screen "Visu_ES_rep5_6" 1280x800, template "Modèle_ES"
   GraphicView "Vue de graphique_1" at 62,186 size 76x151; Picture "Graphique_4"
   TextField "Champ de texte_1" at 43,144 size 59x25; Text 'REP 5'
   Rectangle "Rectangle_2" at 189,244 size 20x20
      Appearance <- "I_det_photo_02"
   TextField "Champ de texte_2" at 215,242 size 136x25; Text 'Det. Photo. 5'
   Rectangle "Rectangle_3" at 189,266 size 20x20
      Appearance <- "AlwaysFALSE"
   TextField "Champ de texte_3" at 215,264 size 53x25; Text 'Libre'
   Rectangle "Rectangle_4" at 189,288 size 20x20
      Appearance <- "AlwaysFALSE"
   TextField "Champ de texte_4" at 215,286 size 53x25; Text 'Libre'
   Rectangle "Rectangle_5" at 189,310 size 20x20
      Appearance <- "AlwaysFALSE"
   TextField "Champ de texte_5" at 215,308 size 53x25; Text 'Libre'
   Rectangle "Rectangle_6" at 189,332 size 20x20
      Appearance <- "AlwaysFALSE"
   TextField "Champ de texte_6" at 215,330 size 53x25; Text 'Libre'
   Rectangle "Rectangle_7" at 189,354 size 20x20
      Appearance <- "AlwaysFALSE"
   TextField "Champ de texte_7" at 215,352 size 53x25; Text 'Libre'
   Rectangle "Rectangle_8" at 189,376 size 20x20
      Appearance <- "AlwaysFALSE"
   TextField "Champ de texte_8" at 215,374 size 53x25; Text 'Libre'
   Rectangle "Rectangle_9" at 189,398 size 20x20
      Appearance <- "AlwaysFALSE"
   TextField "Champ de texte_9" at 215,396 size 53x25; Text 'Libre'
   Rectangle "Rectangle_10" at 399,244 size 20x20
      Appearance <- "I_det_photo_01"
   TextField "Champ de texte_10" at 425,242 size 136x25; Text 'Det. Photo. 4'
   Rectangle "Rectangle_11" at 399,266 size 20x20
      Appearance <- "I_det_photo_03"
   TextField "Champ de texte_11" at 425,264 size 136x25; Text 'Det. Photo. 6'
   Rectangle "Rectangle_12" at 399,288 size 20x20
      Appearance <- "AlwaysFALSE"
   TextField "Champ de texte_12" at 425,286 size 53x25; Text 'Libre'
   Rectangle "Rectangle_13" at 399,310 size 20x20
      Appearance <- "I_libre_I23"
   TextField "Champ de texte_13" at 425,308 size 53x25; Text 'Libre'
   Rectangle "Rectangle_14" at 399,332 size 20x20
      Appearance <- "AlwaysFALSE"
   TextField "Champ de texte_14" at 425,330 size 53x25; Text 'Libre'
   Rectangle "Rectangle_15" at 399,354 size 20x20
      Appearance <- "AlwaysFALSE"
   TextField "Champ de texte_15" at 425,352 size 53x25; Text 'Libre'
   Rectangle "Rectangle_16" at 399,376 size 20x20
      Appearance <- "AlwaysFALSE"
   TextField "Champ de texte_16" at 425,374 size 53x25; Text 'Libre'
   Rectangle "Rectangle_17" at 399,398 size 20x20
      Appearance <- "AlwaysFALSE"
   TextField "Champ de texte_17" at 425,396 size 53x25; Text 'Libre'
   TextField "Champ de texte_34" at 170,173 size 459x25; Text 'ENTREES'
   TextField "Champ de texte_35" at 189,219 size 59x25; Text '%I12'
   TextField "Champ de texte_37" at 399,219 size 59x25; Text '%I13'
   GraphicView "Vue de graphique_2" at 62,454 size 76x151; Picture "Graphique_4"
   TextField "Champ de texte_18" at 43,412 size 59x25; Text 'REP 6'
   Rectangle "Rectangle_20" at 189,512 size 20x20
      Appearance <- "I_Det_Photo_8"
   TextField "Champ de texte_19" at 215,510 size 130x25; Text 'Det. Photo. 8'
   Rectangle "Rectangle_21" at 189,534 size 20x20
      Appearance <- "AlwaysFALSE"
   TextField "Champ de texte_20" at 215,532 size 53x25; Text 'Libre'
   Rectangle "Rectangle_22" at 189,556 size 20x20
      Appearance <- "AlwaysFALSE"
   TextField "Champ de texte_21" at 215,554 size 53x25; Text 'Libre'
   Rectangle "Rectangle_23" at 189,578 size 20x20
      Appearance <- "AlwaysFALSE"
   TextField "Champ de texte_22" at 215,576 size 53x25; Text 'Libre'
   Rectangle "Rectangle_24" at 189,600 size 20x20
      Appearance <- "AlwaysFALSE"
   TextField "Champ de texte_23" at 215,598 size 53x25; Text 'Libre'
   Rectangle "Rectangle_25" at 189,622 size 20x20
      Appearance <- "AlwaysFALSE"
   TextField "Champ de texte_24" at 215,620 size 53x25; Text 'Libre'
   Rectangle "Rectangle_26" at 189,644 size 20x20
      Appearance <- "AlwaysFALSE"
   TextField "Champ de texte_25" at 215,642 size 53x25; Text 'Libre'
   Rectangle "Rectangle_27" at 189,666 size 20x20
      Appearance <- "AlwaysFALSE"
   TextField "Champ de texte_26" at 215,664 size 53x25; Text 'Libre'
   Rectangle "Rectangle_28" at 399,512 size 20x20
      Appearance <- "I_Det_Photo_7"
   TextField "Champ de texte_27" at 425,510 size 130x25; Text 'Det. Photo. 7'
   Rectangle "Rectangle_29" at 399,534 size 20x20
      Appearance <- "I_Det_Photo_9"
   TextField "Champ de texte_28" at 425,532 size 130x25; Text 'Det. Photo. 9'
   Rectangle "Rectangle_30" at 399,556 size 20x20
      Appearance <- "AlwaysFALSE"
   TextField "Champ de texte_29" at 425,554 size 53x25; Text 'Libre'
   Rectangle "Rectangle_31" at 399,578 size 20x20
      Appearance <- "AlwaysFALSE"
   TextField "Champ de texte_30" at 425,576 size 53x25; Text 'Libre'
   Rectangle "Rectangle_32" at 399,600 size 20x20
      Appearance <- "AlwaysFALSE"
   TextField "Champ de texte_31" at 425,598 size 53x25; Text 'Libre'
   Rectangle "Rectangle_34" at 399,622 size 20x20
      Appearance <- "AlwaysFALSE"
   TextField "Champ de texte_32" at 425,620 size 53x25; Text 'Libre'
   Rectangle "Rectangle_36" at 399,644 size 20x20
      Appearance <- "AlwaysFALSE"
   TextField "Champ de texte_33" at 425,642 size 53x25; Text 'Libre'
   Rectangle "Rectangle_37" at 399,666 size 20x20
      Appearance <- "AlwaysFALSE"
   TextField "Champ de texte_36" at 425,664 size 53x25; Text 'Libre'
   TextField "Champ de texte_38" at 170,441 size 459x25; Text 'ENTREES'
   TextField "Champ de texte_39" at 189,487 size 59x25; Text '%I14'
   TextField "Champ de texte_40" at 399,487 size 59x25; Text '%I15'

screen "Visu_ES_Ilot01" 1280x800, template "Modèle_ES"
   TextField "Champ de texte_1" at 43,144 size 80x25; Text 'ILOT 01'
   Rectangle "Rectangle_2" at 273,244 size 20x20
      Appearance <- "O_Rentrer_Butée_01"
   TextField "Champ de texte_2" at 299,242 size 167x25; Text 'Rentrer Butée 01'
   Rectangle "Rectangle_3" at 273,266 size 20x20
      Appearance <- "O_Rentrer_Butée_EL_01"
   TextField "Champ de texte_3" at 299,264 size 202x25; Text 'Rentrer But. Elev. 01'
   Rectangle "Rectangle_4" at 273,288 size 20x20
      Appearance <- "O_Monter_EL_01"
   TextField "Champ de texte_4" at 299,286 size 184x25; Text 'Sortir Elevateur 01'
   Rectangle "Rectangle_5" at 273,310 size 20x20
      Appearance <- "O_Desc_EL_01"
   TextField "Champ de texte_5" at 299,308 size 201x25; Text 'Rentrer Elevateur 01'
   Rectangle "Rectangle_6" at 273,332 size 20x20
      Appearance <- "O_Rentrer_Butée_02"
   TextField "Champ de texte_6" at 299,330 size 167x25; Text 'Rentrer Butée 02'
   Rectangle "Rectangle_7" at 273,354 size 20x20
      Appearance <- "O_Rentrer_Butée_EL_02"
   TextField "Champ de texte_7" at 299,352 size 202x25; Text 'Rentrer But. Elev. 02'
   Rectangle "Rectangle_8" at 273,376 size 20x20
      Appearance <- "O_Monter_EL_02"
   TextField "Champ de texte_8" at 299,374 size 184x25; Text 'Sortir Elevateur 02'
   Rectangle "Rectangle_9" at 273,398 size 20x20
      Appearance <- "O_Desc_EL_02"
   TextField "Champ de texte_9" at 299,396 size 201x25; Text 'Rentrer Elevateur 02'
   Rectangle "Rectangle_10" at 483,244 size 20x20
      Appearance <- "O_Rentrer_Butée_03"
   TextField "Champ de texte_10" at 509,242 size 167x25; Text 'Rentrer Butée 03'
   Rectangle "Rectangle_11" at 483,266 size 20x20
      Appearance <- "O_Rentrer_Butée_EL_03"
   TextField "Champ de texte_11" at 509,264 size 202x25; Text 'Rentrer But. Elev. 03'
   Rectangle "Rectangle_12" at 483,288 size 20x20
      Appearance <- "O_Monter_EL_03"
   TextField "Champ de texte_12" at 509,286 size 184x25; Text 'Sortir Elevateur 03'
   Rectangle "Rectangle_13" at 483,310 size 20x20
      Appearance <- "O_Desc_EL_03"
   TextField "Champ de texte_13" at 509,308 size 201x25; Text 'Rentrer Elevateur 03'
   Rectangle "Rectangle_14" at 483,332 size 20x20
      Appearance <- "O_Rentrer_Butée_04"
   TextField "Champ de texte_14" at 509,330 size 167x25; Text 'Rentrer Butée 04'
   Rectangle "Rectangle_15" at 483,354 size 20x20
      Appearance <- "O_Rentrer_Butée_EL_04"
   TextField "Champ de texte_15" at 509,352 size 202x25; Text 'Rentrer But. Elev. 04'
   Rectangle "Rectangle_16" at 483,376 size 20x20
      Appearance <- "O_Monter_EL_04"
   TextField "Champ de texte_16" at 509,374 size 184x25; Text 'Sortir Elevateur 04'
   Rectangle "Rectangle_17" at 483,398 size 20x20
      Appearance <- "O_Desc_EL_04"
   TextField "Champ de texte_17" at 509,396 size 201x25; Text 'Rentrer Elevateur 04'
   TextField "Champ de texte_34" at 254,173 size 880x25; Text 'SORTIES'
   TextField "Champ de texte_35" at 273,219 size 64x25; Text '%Q10'
   TextField "Champ de texte_37" at 483,219 size 64x25; Text '%Q11'
   GraphicView "Vue de graphique_3" at 58,184 size 154x109; Picture "Graphique_5"
   Rectangle "Rectangle_18" at 692,244 size 20x20
      Appearance <- "O_Rentrer_Butée_05"
   TextField "Champ de texte_18" at 718,242 size 167x25; Text 'Rentrer Butée 05'
   Rectangle "Rectangle_19" at 692,266 size 20x20
      Appearance <- "O_Rentrer_Butée_EL_05"
   TextField "Champ de texte_19" at 718,264 size 202x25; Text 'Rentrer But. Elev. 05'
   Rectangle "Rectangle_20" at 692,288 size 20x20
      Appearance <- "O_Monter_EL_05"
   TextField "Champ de texte_20" at 718,286 size 184x25; Text 'Sortir Elevateur 05'
   Rectangle "Rectangle_21" at 692,310 size 20x20
      Appearance <- "O_Desc_EL_05"
   TextField "Champ de texte_21" at 718,308 size 201x25; Text 'Rentrer Elevateur 05'
   Rectangle "Rectangle_22" at 692,332 size 20x20
      Appearance <- "O_Rentrer_Butée_06"
   TextField "Champ de texte_22" at 718,330 size 167x25; Text 'Rentrer Butée 06'
   Rectangle "Rectangle_23" at 692,354 size 20x20
      Appearance <- "O_Rentrer_Butée_EL_06"
   TextField "Champ de texte_23" at 718,352 size 202x25; Text 'Rentrer But. Elev. 06'
   Rectangle "Rectangle_24" at 692,376 size 20x20
      Appearance <- "O_Monter_EL_06"
   TextField "Champ de texte_24" at 718,374 size 184x25; Text 'Sortir Elevateur 06'
   Rectangle "Rectangle_25" at 692,398 size 20x20
      Appearance <- "O_Desc_EL_06"
   TextField "Champ de texte_25" at 718,396 size 201x25; Text 'Rentrer Elevateur 06'
   Rectangle "Rectangle_26" at 902,244 size 20x20
      Appearance <- "O_Rentrer_Butée_07"
   TextField "Champ de texte_26" at 928,242 size 167x25; Text 'Rentrer Butée 07'
   Rectangle "Rectangle_27" at 902,266 size 20x20
      Appearance <- "O_Rentrer_Butée_EL_07"
   TextField "Champ de texte_27" at 928,264 size 202x25; Text 'Rentrer But. Elev. 07'
   Rectangle "Rectangle_28" at 902,288 size 20x20
      Appearance <- "O_Monter_EL_07"
   TextField "Champ de texte_28" at 928,286 size 184x25; Text 'Sortir Elevateur 07'
   Rectangle "Rectangle_29" at 902,310 size 20x20
      Appearance <- "O_Desc_EL_07"
   TextField "Champ de texte_29" at 928,308 size 201x25; Text 'Rentrer Elevateur 07'
   Rectangle "Rectangle_30" at 902,332 size 20x20
      Appearance <- "O_Op_Porte_Vision"
   TextField "Champ de texte_30" at 928,330 size 185x25; Text 'Ouvrir Porte Vision'
   Rectangle "Rectangle_31" at 902,354 size 20x20
      Appearance <- "O_Cl_porte_Vision"
   TextField "Champ de texte_31" at 928,352 size 192x25; Text 'Fermer Porte Vision'
   Rectangle "Rectangle_32" at 902,376 size 20x20
      Appearance <- "I_libre_I26"
   TextField "Champ de texte_32" at 928,374 size 53x25; Text 'Libre'
   Rectangle "Rectangle_34" at 902,398 size 20x20
      Appearance <- "I_libre_I27"
   TextField "Champ de texte_33" at 928,396 size 53x25; Text 'Libre'
   TextField "Champ de texte_36" at 692,219 size 64x25; Text '%Q12'
   TextField "Champ de texte_38" at 902,219 size 64x25; Text '%Q13'

screen "Visu_ES_Ilot02" 1280x800, template "Modèle_ES"
   TextField "Champ de texte_1" at 43,144 size 80x25; Text 'ILOT 02'
   Rectangle "Rectangle_2" at 273,244 size 20x20
      Appearance <- "O_Sortir_Blocage_boite_01"
   TextField "Champ de texte_2" at 299,242 size 184x25; Text 'Sortir Verin 1 bloc.'
   Rectangle "Rectangle_3" at 273,266 size 20x20
      Appearance <- "O_Rentrer_Blocage_boite_01"
   TextField "Champ de texte_3" at 299,264 size 201x25; Text 'Rentrer Verin 1 bloc.'
   Rectangle "Rectangle_4" at 273,288 size 20x20
      Appearance <- "O_Sortir_Blocage_boite_02"
   TextField "Champ de texte_4" at 299,286 size 184x25; Text 'Sortir Verin 2 bloc.'
   Rectangle "Rectangle_5" at 273,310 size 20x20
      Appearance <- "O_Rentrer_Blocage_boite_02"
   TextField "Champ de texte_5" at 299,308 size 201x25; Text 'Rentrer Verin 2 bloc.'
   Rectangle "Rectangle_6" at 273,332 size 20x20
      Appearance <- "O_Sortir_Blocage_boite_03"
   TextField "Champ de texte_6" at 299,330 size 184x25; Text 'Sortir Verin 3 bloc.'
   Rectangle "Rectangle_7" at 273,354 size 20x20
      Appearance <- "O_Rentrer_Blocage_boite_03"
   TextField "Champ de texte_7" at 299,352 size 201x25; Text 'Rentrer Verin 3 bloc.'
   Rectangle "Rectangle_8" at 273,376 size 20x20
      Appearance <- "O_Sortir_Blocage_boite_04"
   TextField "Champ de texte_8" at 299,374 size 184x25; Text 'Sortir Verin 4 bloc.'
   Rectangle "Rectangle_9" at 273,398 size 20x20
      Appearance <- "O_Rentrer_Blocage_boite_04"
   TextField "Champ de texte_9" at 299,396 size 201x25; Text 'Rentrer Verin 4 bloc.'
   Rectangle "Rectangle_10" at 483,244 size 20x20
      Appearance <- "I_libre_I20"
   TextField "Champ de texte_10" at 509,242 size 53x25; Text 'Libre'
   Rectangle "Rectangle_11" at 483,266 size 20x20
      Appearance <- "I_libre_I21"
   TextField "Champ de texte_11" at 509,264 size 53x25; Text 'Libre'
   Rectangle "Rectangle_12" at 483,288 size 20x20
      Appearance <- "I_libre_I22"
   TextField "Champ de texte_12" at 509,286 size 53x25; Text 'Libre'
   Rectangle "Rectangle_13" at 483,310 size 20x20
      Appearance <- "I_libre_I23"
   TextField "Champ de texte_13" at 509,308 size 53x25; Text 'Libre'
   Rectangle "Rectangle_14" at 483,332 size 20x20
      Appearance <- "I_libre_I24"
   TextField "Champ de texte_14" at 509,330 size 53x25; Text 'Libre'
   Rectangle "Rectangle_15" at 483,354 size 20x20
      Appearance <- "I_libre_I25"
   TextField "Champ de texte_15" at 509,352 size 53x25; Text 'Libre'
   Rectangle "Rectangle_16" at 483,376 size 20x20
      Appearance <- "I_libre_I26"
   TextField "Champ de texte_16" at 509,374 size 53x25; Text 'Libre'
   Rectangle "Rectangle_17" at 483,398 size 20x20
      Appearance <- "I_libre_I27"
   TextField "Champ de texte_17" at 509,396 size 53x25; Text 'Libre'
   TextField "Champ de texte_34" at 254,173 size 880x25; Text 'SORTIES'
   TextField "Champ de texte_35" at 273,219 size 64x25; Text '%Q14'
   TextField "Champ de texte_37" at 483,219 size 64x25; Text '%Q15'
   GraphicView "Vue de graphique_3" at 58,184 size 154x109; Picture "Graphique_5"
   Rectangle "Rectangle_18" at 692,244 size 20x20
      Appearance <- "I_En_Service"
   TextField "Champ de texte_18" at 718,242 size 53x25; Text 'Libre'
   Rectangle "Rectangle_19" at 692,266 size 20x20
      Appearance <- "I_En_Arret_Urgence"
   TextField "Champ de texte_19" at 718,264 size 53x25; Text 'Libre'
   Rectangle "Rectangle_20" at 692,288 size 20x20
      Appearance <- "I_En_Manuel"
   TextField "Champ de texte_20" at 718,286 size 53x25; Text 'Libre'
   Rectangle "Rectangle_21" at 692,310 size 20x20
      Appearance <- "I_En_Automatique"
   TextField "Champ de texte_21" at 718,308 size 53x25; Text 'Libre'
   Rectangle "Rectangle_22" at 692,332 size 20x20
      Appearance <- "I_porte_non_réarmée"
   TextField "Champ de texte_22" at 718,330 size 53x25; Text 'Libre'
   Rectangle "Rectangle_23" at 692,354 size 20x20
      Appearance <- "I_porte_01_Op"
   TextField "Champ de texte_23" at 718,352 size 53x25; Text 'Libre'
   Rectangle "Rectangle_24" at 692,376 size 20x20
      Appearance <- "I_porte_02_Op"
   TextField "Champ de texte_24" at 718,374 size 53x25; Text 'Libre'
   Rectangle "Rectangle_25" at 692,398 size 20x20
      Appearance <- "I_libre_I07"
   TextField "Champ de texte_25" at 718,396 size 53x25; Text 'Libre'
   Rectangle "Rectangle_26" at 902,244 size 20x20
      Appearance <- "I_libre_I20"
   TextField "Champ de texte_26" at 928,242 size 53x25; Text 'Libre'
   Rectangle "Rectangle_27" at 902,266 size 20x20
      Appearance <- "I_libre_I21"
   TextField "Champ de texte_27" at 928,264 size 53x25; Text 'Libre'
   Rectangle "Rectangle_28" at 902,288 size 20x20
      Appearance <- "I_libre_I22"
   TextField "Champ de texte_28" at 928,286 size 53x25; Text 'Libre'
   Rectangle "Rectangle_29" at 902,310 size 20x20
      Appearance <- "I_libre_I23"
   TextField "Champ de texte_29" at 928,308 size 53x25; Text 'Libre'
   Rectangle "Rectangle_30" at 902,332 size 20x20
      Appearance <- "I_libre_I24"
   TextField "Champ de texte_30" at 928,330 size 53x25; Text 'Libre'
   Rectangle "Rectangle_31" at 902,354 size 20x20
      Appearance <- "I_libre_I25"
   TextField "Champ de texte_31" at 928,352 size 53x25; Text 'Libre'
   Rectangle "Rectangle_32" at 902,376 size 20x20
      Appearance <- "I_libre_I26"
   TextField "Champ de texte_32" at 928,374 size 53x25; Text 'Libre'
   Rectangle "Rectangle_34" at 902,398 size 20x20
      Appearance <- "I_libre_I27"
   TextField "Champ de texte_33" at 928,396 size 53x25; Text 'Libre'
   TextField "Champ de texte_36" at 692,219 size 64x25; Text '%Q16'
   TextField "Champ de texte_38" at 902,219 size 64x25; Text '%Q17'

screen "Mode_Manuel_B01" 1280x800, template "Modèle_Manu"
   TextField "Champ de texte_34" at 33,135 size 584x25; Text 'Hyppodrome Poste 01'
   Button "Bouton_1" at 39,179 size 169x68; TextOff 'MONTER BUTEE'
      on Press: SetBit("Touche_Tch_Manu{0}")
      on Release: ResetBit("Touche_Tch_Manu{0}")
      Appearance <- "O_Rentrer_Butée_01"
   Button "Bouton_2" at 39,255 size 169x68; TextOff 'DESCENDRE BUTEE'
      on Press: SetBit("Touche_Tch_Manu{1}")
      on Release: ResetBit("Touche_Tch_Manu{1}")
   Button "Bouton_3" at 220,179 size 169x68; TextOff 'MONTER BUTEE ELEVATEUR'
      on Press: SetBit("Touche_Tch_Manu{2}")
      on Release: ResetBit("Touche_Tch_Manu{2}")
   Button "Bouton_4" at 220,255 size 169x68; TextOff 'DESCENDRE BUTEE ELEVATEUR'
      on Press: SetBit("Touche_Tch_Manu{3}")
      on Release: ResetBit("Touche_Tch_Manu{3}")
   Button "Bouton_5" at 39,331 size 169x68; TextOff 'MONTER ELEVATEUR'
      on Press: SetBit("Touche_Tch_Manu{4}")
      on Release: ResetBit("Touche_Tch_Manu{4}")
   Button "Bouton_6" at 220,331 size 169x68; TextOff 'DESCENDRE ELEVATEUR'
      on Press: SetBit("Touche_Tch_Manu{5}")
      on Release: ResetBit("Touche_Tch_Manu{5}")
   Rectangle "Rectangle_2" at 404,181 size 20x20
      Appearance <- "I_Pres_Pal_B01"
   TextField "Champ de texte_2" at 430,179 size 168x25; Text 'Presence pal B01'
   Rectangle "Rectangle_3" at 404,203 size 20x20
      Appearance <- "I_Pres_Elev_B01"
   TextField "Champ de texte_3" at 430,201 size 178x25; Text 'Presence Elev B01'
   Rectangle "Rectangle_4" at 404,225 size 20x20
      Appearance <- "I_Elev_01_Bas"
   TextField "Champ de texte_4" at 430,223 size 177x25; Text 'Elevateur Bas B01'
   Rectangle "Rectangle_5" at 404,247 size 20x20
      Appearance <- "I_Elev_01_Haut"
   TextField "Champ de texte_5" at 430,245 size 188x25; Text 'Elevateur Haut B01'
   TextField "Champ de texte_1" at 34,419 size 584x25; Text 'Hyppodrome Poste 02'
   Button "Bouton_7" at 38,460 size 169x68; TextOff 'MONTER BUTEE'
      on Release: ResetBit("Touche_Tch_Manu{6}")
      on Press: SetBit("Touche_Tch_Manu{6}")
   Button "Bouton_8" at 38,536 size 169x68; TextOff 'DESCENDRE BUTEE'
      on Release: ResetBit("Touche_Tch_Manu{7}")
      on Press: SetBit("Touche_Tch_Manu{7}")
   Button "Bouton_9" at 219,460 size 169x68; TextOff 'MONTER BUTEE ELEVATEUR'
      on Release: ResetBit("Touche_Tch_Manu{8}")
      on Press: SetBit("Touche_Tch_Manu{8}")
   Button "Bouton_10" at 219,536 size 169x68; TextOff 'DESCENDRE BUTEE ELEVATEUR'
      on Release: ResetBit("Touche_Tch_Manu{9}")
      on Press: SetBit("Touche_Tch_Manu{9}")
   Button "Bouton_11" at 38,612 size 169x68; TextOff 'MONTER ELEVATEUR'
      on Release: ResetBit("Touche_Tch_Manu{10}")
      on Press: SetBit("Touche_Tch_Manu{10}")
   Button "Bouton_12" at 219,612 size 169x68; TextOff 'DESCENDRE ELEVATEUR'
      on Release: ResetBit("Touche_Tch_Manu{11}")
      on Press: SetBit("Touche_Tch_Manu{11}")
   Rectangle "Rectangle_7" at 403,462 size 20x20
      Appearance <- "I_Pres_Pal_B02"
   TextField "Champ de texte_6" at 429,460 size 168x25; Text 'Presence pal B02'
   Rectangle "Rectangle_8" at 403,484 size 20x20
      Appearance <- "I_Pres_Elev_B02"
   TextField "Champ de texte_7" at 429,482 size 178x25; Text 'Presence Elev B02'
   Rectangle "Rectangle_9" at 403,506 size 20x20
      Appearance <- "I_Elev_02_Bas"
   TextField "Champ de texte_8" at 429,504 size 177x25; Text 'Elevateur Bas B02'
   Rectangle "Rectangle_10" at 403,528 size 20x20
      Appearance <- "I_Elev_02_Haut"
   TextField "Champ de texte_9" at 429,526 size 188x25; Text 'Elevateur Haut B02'
   TextField "Champ de texte_10" at 665,138 size 584x25; Text 'Hyppodrome Poste 03'
   Button "Bouton_13" at 669,179 size 169x68; TextOff 'MONTER BUTEE'
      on Release: ResetBit("Touche_Tch_Manu{12}")
      on Press: SetBit("Touche_Tch_Manu{12}")
   Button "Bouton_14" at 669,255 size 169x68; TextOff 'DESCENDRE BUTEE'
      on Release: ResetBit("Touche_Tch_Manu{13}")
      on Press: SetBit("Touche_Tch_Manu{13}")
   Button "Bouton_15" at 850,179 size 169x68; TextOff 'MONTER BUTEE ELEVATEUR'
      on Release: ResetBit("Touche_Tch_Manu{14}")
      on Press: SetBit("Touche_Tch_Manu{14}")
   Button "Bouton_16" at 850,255 size 169x68; TextOff 'DESCENDRE BUTEE ELEVATEUR'
      on Release: ResetBit("Touche_Tch_Manu{15}")
      on Press: SetBit("Touche_Tch_Manu{15}")
   Button "Bouton_17" at 669,331 size 169x68; TextOff 'MONTER ELEVATEUR'
      on Release: ResetBit("Touche_Tch_Manu{16}")
      on Press: SetBit("Touche_Tch_Manu{16}")
   Button "Bouton_18" at 850,331 size 169x68; TextOff 'DESCENDRE ELEVATEUR'
      on Release: ResetBit("Touche_Tch_Manu{17}")
      on Press: SetBit("Touche_Tch_Manu{17}")
   Rectangle "Rectangle_13" at 1034,181 size 20x20
      Appearance <- "I_Pres_Pal_B03"
   TextField "Champ de texte_11" at 1060,179 size 168x25; Text 'Presence pal B03'
   Rectangle "Rectangle_14" at 1034,203 size 20x20
      Appearance <- "I_Pres_Elev_B03"
   TextField "Champ de texte_12" at 1060,201 size 178x25; Text 'Presence Elev B03'
   Rectangle "Rectangle_15" at 1034,225 size 20x20
      Appearance <- "I_Elev_03_Bas"
   TextField "Champ de texte_13" at 1060,223 size 177x25; Text 'Elevateur Bas B03'
   Rectangle "Rectangle_16" at 1034,247 size 20x20
      Appearance <- "I_Elev_03_Haut"
   TextField "Champ de texte_14" at 1060,245 size 188x25; Text 'Elevateur Haut B03'
   TextField "Champ de texte_15" at 664,419 size 584x25; Text 'Hyppodrome Poste 04'
   Button "Bouton_19" at 668,460 size 169x68; TextOff 'MONTER BUTEE'
      on Release: ResetBit("Touche_Tch_Manu{18}")
      on Press: SetBit("Touche_Tch_Manu{18}")
   Button "Bouton_20" at 668,536 size 169x68; TextOff 'DESCENDRE BUTEE'
      on Release: ResetBit("Touche_Tch_Manu{19}")
      on Press: SetBit("Touche_Tch_Manu{19}")
   Button "Bouton_21" at 849,460 size 169x68; TextOff 'MONTER BUTEE ELEVATEUR'
      on Release: ResetBit("Touche_Tch_Manu{20}")
      on Press: SetBit("Touche_Tch_Manu{20}")
   Button "Bouton_22" at 849,536 size 169x68; TextOff 'DESCENDRE BUTEE ELEVATEUR'
      on Release: ResetBit("Touche_Tch_Manu{21}")
      on Press: SetBit("Touche_Tch_Manu{21}")
   Button "Bouton_23" at 668,612 size 169x68; TextOff 'MONTER ELEVATEUR'
      on Release: ResetBit("Touche_Tch_Manu{22}")
      on Press: SetBit("Touche_Tch_Manu{22}")
   Button "Bouton_24" at 849,612 size 169x68; TextOff 'DESCENDRE ELEVATEUR'
      on Release: ResetBit("Touche_Tch_Manu{23}")
      on Press: SetBit("Touche_Tch_Manu{23}")
   Rectangle "Rectangle_19" at 1033,462 size 20x20
      Appearance <- "I_Pres_Pal_B04"
   TextField "Champ de texte_16" at 1059,460 size 168x25; Text 'Presence pal B04'
   Rectangle "Rectangle_20" at 1033,484 size 20x20
      Appearance <- "I_Pres_Elev_B04"
   TextField "Champ de texte_17" at 1059,482 size 178x25; Text 'Presence Elev B04'
   Rectangle "Rectangle_21" at 1033,506 size 20x20
      Appearance <- "I_Elev_04_Bas"
   TextField "Champ de texte_18" at 1059,504 size 177x25; Text 'Elevateur Bas B04'
   Rectangle "Rectangle_22" at 1033,528 size 20x20
      Appearance <- "I_Elev_04_Haut"
   TextField "Champ de texte_19" at 1059,526 size 188x25; Text 'Elevateur Haut B04'
   Rectangle "Rectangle_23" at 404,285 size 20x20
      Appearance <- "O_Rentrer_Butée_01"
   TextField "Champ de texte_20" at 430,283 size 137x25; Text 'Rentrer Butée'
   Rectangle "Rectangle_24" at 404,307 size 20x20
      Appearance <- "O_Rentrer_Butée_EL_01"
   TextField "Champ de texte_21" at 430,305 size 188x25; Text 'Rentrer Butée Elev.'
   Rectangle "Rectangle_25" at 404,329 size 20x20
      Appearance <- "O_Monter_EL_01"
   TextField "Champ de texte_22" at 430,327 size 167x25; Text 'Monter Elevateur'
   Rectangle "Rectangle_26" at 404,351 size 20x20
      Appearance <- "O_Desc_EL_01"
   TextField "Champ de texte_23" at 430,349 size 199x25; Text 'Descendre Elevateur'
   Rectangle "Rectangle_27" at 1034,287 size 20x20
      Appearance <- "O_Rentrer_Butée_03"
   TextField "Champ de texte_24" at 1060,285 size 137x25; Text 'Rentrer Butée'
   Rectangle "Rectangle_28" at 1034,309 size 20x20
      Appearance <- "O_Rentrer_Butée_EL_03"
   TextField "Champ de texte_25" at 1060,307 size 188x25; Text 'Rentrer Butée Elev.'
   Rectangle "Rectangle_29" at 1034,331 size 20x20
      Appearance <- "O_Monter_EL_03"
   TextField "Champ de texte_26" at 1060,329 size 167x25; Text 'Monter Elevateur'
   Rectangle "Rectangle_30" at 1034,353 size 20x20
      Appearance <- "O_Desc_EL_03"
   TextField "Champ de texte_27" at 1060,351 size 199x25; Text 'Descendre Elevateur'
   Rectangle "Rectangle_31" at 403,571 size 20x20
      Appearance <- "O_Rentrer_Butée_02"
   TextField "Champ de texte_28" at 429,569 size 137x25; Text 'Rentrer Butée'
   Rectangle "Rectangle_32" at 403,593 size 20x20
      Appearance <- "O_Rentrer_Butée_EL_02"
   TextField "Champ de texte_29" at 429,591 size 188x25; Text 'Rentrer Butée Elev.'
   Rectangle "Rectangle_34" at 403,615 size 20x20
      Appearance <- "O_Monter_EL_02"
   TextField "Champ de texte_30" at 429,613 size 167x25; Text 'Monter Elevateur'
   Rectangle "Rectangle_36" at 403,637 size 20x20
      Appearance <- "O_Desc_EL_02"
   TextField "Champ de texte_31" at 429,635 size 199x25; Text 'Descendre Elevateur'
   Rectangle "Rectangle_37" at 1034,573 size 20x20
      Appearance <- "O_Rentrer_Butée_04"
   TextField "Champ de texte_32" at 1060,571 size 137x25; Text 'Rentrer Butée'
   Rectangle "Rectangle_38" at 1034,595 size 20x20
      Appearance <- "O_Rentrer_Butée_EL_04"
   TextField "Champ de texte_33" at 1060,593 size 188x25; Text 'Rentrer Butée Elev.'
   Rectangle "Rectangle_39" at 1034,617 size 20x20
      Appearance <- "O_Monter_EL_04"
   TextField "Champ de texte_35" at 1060,615 size 167x25; Text 'Monter Elevateur'
   Rectangle "Rectangle_40" at 1034,639 size 20x20
      Appearance <- "O_Desc_EL_04"
   TextField "Champ de texte_36" at 1059,637 size 199x25; Text 'Descendre Elevateur'

Template "Modèle_Manu" 1280x800
   Button "Bouton_1" at 968,723 size 96x70; TextOff 'Text'
   Button "Bouton_5" at 861,723 size 96x70; TextOff 'Imp 3D'
      on Release: ActivateScreen("Mode_Manuel_Imprimantes", 0)
   Button "Bouton_6" at 754,723 size 96x70; TextOff 'Vision'
      on Release: ActivateScreen("Mode_Manuel_Vision", 0)
      ObjectEnable <- "Bits_Globaux_x_En_manu"
   Button "Bouton_7" at 647,723 size 96x70; TextOff 'CONV. CART. 03'
      on Release: ActivateScreen("Mode_Manuel_Conv_carton_03", 0)
      ObjectEnable <- "Bits_Globaux_x_En_manu"
   Button "Bouton_8" at 540,723 size 96x70; TextOff 'CONV. CART. 02'
      on Release: ActivateScreen("Mode_Manuel_Conv_carton_02", 0)
      ObjectEnable <- "Bits_Globaux_x_En_manu"
   Button "Bouton_9" at 433,723 size 96x70; TextOff 'CONV. CART. 01'
      on Release: ActivateScreen("Mode_Manuel_Conv_carton_01", 0)
      ObjectEnable <- "Bits_Globaux_x_En_manu"
   Button "Bouton_10" at 326,723 size 96x70; TextOff 'VERIN BLOCAGE'
      on Release: ActivateScreen("Mode_Manuel_Conv_carton", 0)
      ObjectEnable <- "Bits_Globaux_x_En_manu"
   Button "Bouton_11" at 219,723 size 96x70; TextOff 'HYPPO. CONV.'
      on Release: ActivateScreen("Mode_Manuel_Conv_H", 0)
      ObjectEnable <- "Bits_Globaux_x_En_manu"
   Button "Bouton_12" at 112,723 size 96x70; TextOff 'HYPPO. B05..B08'
      on Release: ActivateScreen("Mode_Manuel_B01_std_2", 0)
      ObjectEnable <- "Bits_Globaux_x_En_manu"
   Button "Bouton_13" at 5,723 size 96x70; TextOff 'HYPPO. B01..B04'
      on Release: ActivateScreen("Mode_Manuel_B01_std_1", 0)
      ObjectEnable <- "Bits_Globaux_x_En_manu"
   Button "Bouton_3" at 1177,723 size 96x70; TextOff 'RETOUR'
      on Release: ActivateScreen("Principale", 0)
   DateTimeField "Champ de date/heure_1" at 1133,29 size 131x34
   DateTimeField "Champ de date/heure_2" at 1152,65 size 99x34
   GraphicView "Vue de graphique_1" at 129,8 size 113x116; Picture "Ascodero"
   TextField "Champ de texte_5" at 634,54 size 173x28; Text 'Usine Ecole 4.0'
   GraphicView "Vue de graphique_2" at 9,8 size 111x116; Picture "unilasalle"
   Button "Bouton_14" at 4,5 size 124x122; TextOff 'Text'
      on Click: ActivateScreen("Page_demarrage", 0)

screen "Mode_Manuel_B02" 1280x800, template "Modèle_Manu"
   TextField "Champ de texte_34" at 35,138 size 584x25; Text 'Hyppodrome Poste 05'
   Button "Bouton_1" at 39,179 size 169x68; TextOff 'MONTER BUTEE'
      on Release: ResetBit("Touche_Tch_Manu{24}")
      on Press: SetBit("Touche_Tch_Manu{24}")
   Button "Bouton_2" at 39,255 size 169x68; TextOff 'DESCENDRE BUTEE'
      on Release: ResetBit("Touche_Tch_Manu{25}")
      on Press: SetBit("Touche_Tch_Manu{25}")
   Button "Bouton_3" at 220,179 size 169x68; TextOff 'MONTER BUTEE ELEVATEUR'
      on Release: ResetBit("Touche_Tch_Manu{26}")
      on Press: SetBit("Touche_Tch_Manu{26}")
   Button "Bouton_4" at 220,255 size 169x68; TextOff 'DESCENDRE BUTEE ELEVATEUR'
      on Release: ResetBit("Touche_Tch_Manu{27}")
      on Press: SetBit("Touche_Tch_Manu{27}")
   Button "Bouton_5" at 39,329 size 169x68; TextOff 'MONTER ELEVATEUR'
      on Release: ResetBit("Touche_Tch_Manu{28}")
      on Press: SetBit("Touche_Tch_Manu{28}")
   Button "Bouton_6" at 220,331 size 169x68; TextOff 'DESCENDRE ELEVATEUR'
      on Release: ResetBit("Touche_Tch_Manu{29}")
      on Press: SetBit("Touche_Tch_Manu{29}")
   Rectangle "Rectangle_2" at 404,181 size 20x20
      Appearance <- "I_Pres_Pal_B05"
   TextField "Champ de texte_2" at 430,179 size 168x25; Text 'Presence pal B05'
   Rectangle "Rectangle_3" at 404,203 size 20x20
      Appearance <- "I_Pres_Elev_B05"
   TextField "Champ de texte_3" at 430,201 size 178x25; Text 'Presence Elev B05'
   Rectangle "Rectangle_4" at 404,225 size 20x20
      Appearance <- "I_Elev_05_Bas"
   TextField "Champ de texte_4" at 430,223 size 177x25; Text 'Elevateur Bas B05'
   Rectangle "Rectangle_5" at 404,247 size 20x20
      Appearance <- "I_Elev_05_Haut"
   TextField "Champ de texte_5" at 430,245 size 188x25; Text 'Elevateur Haut B05'
   TextField "Champ de texte_1" at 34,419 size 584x25; Text 'Hyppodrome Poste 06'
   Button "Bouton_7" at 38,460 size 169x68; TextOff 'MONTER BUTEE'
      on Release: ResetBit("Touche_Tch_Manu{30}")
      on Press: SetBit("Touche_Tch_Manu{30}")
   Button "Bouton_8" at 38,536 size 169x68; TextOff 'DESCENDRE BUTEE'
      on Release: ResetBit("Touche_Tch_Manu{31}")
      on Press: SetBit("Touche_Tch_Manu{31}")
   Button "Bouton_9" at 219,460 size 169x68; TextOff 'MONTER BUTEE ELEVATEUR'
      on Release: ResetBit("Touche_Tch_Manu{32}")
      on Press: SetBit("Touche_Tch_Manu{32}")
   Button "Bouton_10" at 219,536 size 169x68; TextOff 'DESCENDRE BUTEE ELEVATEUR'
      on Release: ResetBit("Touche_Tch_Manu{33}")
      on Press: SetBit("Touche_Tch_Manu{33}")
   Button "Bouton_11" at 38,610 size 169x68; TextOff 'MONTER ELEVATEUR'
      on Release: ResetBit("Touche_Tch_Manu{34}")
      on Press: SetBit("Touche_Tch_Manu{34}")
   Button "Bouton_12" at 219,612 size 169x68; TextOff 'DESCENDRE ELEVATEUR'
      on Release: ResetBit("Touche_Tch_Manu{35}")
      on Press: SetBit("Touche_Tch_Manu{35}")
   Rectangle "Rectangle_7" at 403,462 size 20x20
      Appearance <- "I_Pres_Pal_B06"
   TextField "Champ de texte_6" at 429,460 size 168x25; Text 'Presence pal B06'
   Rectangle "Rectangle_8" at 403,484 size 20x20
      Appearance <- "I_Pres_Elev_B06"
   TextField "Champ de texte_7" at 429,482 size 178x25; Text 'Presence Elev B06'
   Rectangle "Rectangle_9" at 403,506 size 20x20
      Appearance <- "I_Elev_06_Bas"
   TextField "Champ de texte_8" at 429,504 size 177x25; Text 'Elevateur Bas B06'
   Rectangle "Rectangle_10" at 403,528 size 20x20
      Appearance <- "I_Elev_06_Haut"
   TextField "Champ de texte_9" at 429,526 size 188x25; Text 'Elevateur Haut B06'
   TextField "Champ de texte_10" at 665,138 size 584x25; Text 'Hyppodrome Poste 07'
   Button "Bouton_13" at 669,179 size 169x68; TextOff 'MONTER BUTEE'
      on Release: ResetBit("Touche_Tch_Manu{36}")
      on Press: SetBit("Touche_Tch_Manu{36}")
   Button "Bouton_14" at 669,255 size 169x68; TextOff 'DESCENDRE BUTEE'
      on Release: ResetBit("Touche_Tch_Manu{37}")
      on Press: SetBit("Touche_Tch_Manu{37}")
   Button "Bouton_15" at 850,179 size 169x68; TextOff 'MONTER BUTEE ELEVATEUR'
      on Release: ResetBit("Touche_Tch_Manu{38}")
      on Press: SetBit("Touche_Tch_Manu{38}")
   Button "Bouton_16" at 850,255 size 169x68; TextOff 'DESCENDRE BUTEE ELEVATEUR'
      on Release: ResetBit("Touche_Tch_Manu{39}")
      on Press: SetBit("Touche_Tch_Manu{39}")
   Button "Bouton_17" at 669,329 size 169x68; TextOff 'MONTER ELEVATEUR'
      on Release: ResetBit("Touche_Tch_Manu{40}")
      on Press: SetBit("Touche_Tch_Manu{40}")
   Button "Bouton_18" at 850,331 size 169x68; TextOff 'DESCENDRE ELEVATEUR'
      on Release: ResetBit("Touche_Tch_Manu{41}")
      on Press: SetBit("Touche_Tch_Manu{41}")
   Rectangle "Rectangle_13" at 1034,181 size 20x20
      Appearance <- "I_Pres_Pal_B07"
   TextField "Champ de texte_11" at 1060,179 size 168x25; Text 'Presence pal B07'
   Rectangle "Rectangle_14" at 1034,203 size 20x20
      Appearance <- "I_Pres_Elev_B07"
   TextField "Champ de texte_12" at 1060,201 size 178x25; Text 'Presence Elev B07'
   Rectangle "Rectangle_15" at 1034,225 size 20x20
      Appearance <- "I_Elev_07_Bas"
   TextField "Champ de texte_13" at 1060,223 size 177x25; Text 'Elevateur Bas B07'
   Rectangle "Rectangle_16" at 1034,247 size 20x20
      Appearance <- "I_Elev_07_Haut"
   TextField "Champ de texte_14" at 1060,245 size 188x25; Text 'Elevateur Haut B07'
   Rectangle "Rectangle_23" at 404,285 size 20x20
      Appearance <- "O_Rentrer_Butée_05"
   TextField "Champ de texte_20" at 430,283 size 137x25; Text 'Rentrer Butée'
   Rectangle "Rectangle_24" at 404,307 size 20x20
      Appearance <- "O_Rentrer_Butée_EL_05"
   TextField "Champ de texte_21" at 430,305 size 188x25; Text 'Rentrer Butée Elev.'
   Rectangle "Rectangle_25" at 404,329 size 20x20
      Appearance <- "O_Monter_EL_05"
   TextField "Champ de texte_22" at 430,327 size 167x25; Text 'Monter Elevateur'
   Rectangle "Rectangle_26" at 404,351 size 20x20
      Appearance <- "O_Desc_EL_05"
   TextField "Champ de texte_23" at 430,349 size 199x25; Text 'Descendre Elevateur'
   Rectangle "Rectangle_31" at 403,571 size 20x20
      Appearance <- "O_Rentrer_Butée_06"
   TextField "Champ de texte_28" at 429,569 size 137x25; Text 'Rentrer Butée'
   Rectangle "Rectangle_32" at 403,593 size 20x20
      Appearance <- "O_Rentrer_Butée_EL_06"
   TextField "Champ de texte_29" at 429,591 size 188x25; Text 'Rentrer Butée Elev.'
   Rectangle "Rectangle_34" at 403,615 size 20x20
      Appearance <- "O_Monter_EL_06"
   TextField "Champ de texte_30" at 429,613 size 167x25; Text 'Monter Elevateur'
   Rectangle "Rectangle_36" at 403,637 size 20x20
      Appearance <- "O_Desc_EL_06"
   TextField "Champ de texte_31" at 429,635 size 199x25; Text 'Descendre Elevateur'
   Rectangle "Rectangle_27" at 1034,287 size 20x20
      Appearance <- "O_Rentrer_Butée_07"
   TextField "Champ de texte_24" at 1060,285 size 137x25; Text 'Rentrer Butée'
   Rectangle "Rectangle_28" at 1034,309 size 20x20
      Appearance <- "O_Rentrer_Butée_EL_07"
   TextField "Champ de texte_25" at 1060,307 size 188x25; Text 'Rentrer Butée Elev.'
   Rectangle "Rectangle_29" at 1034,331 size 20x20
      Appearance <- "O_Monter_EL_07"
   TextField "Champ de texte_26" at 1060,329 size 167x25; Text 'Monter Elevateur'
   Rectangle "Rectangle_30" at 1034,353 size 20x20
      Appearance <- "O_Desc_EL_07"
   TextField "Champ de texte_27" at 1060,351 size 199x25; Text 'Descendre Elevateur'
   Group "Group" at 661,416 size 591x157
   TextField "Champ de texte_15" at 665,419 size 584x25; Text 'Porte Poste Vision'
   Button "Bouton_19" at 669,460 size 169x68; TextOff 'OUVRIR PORTE'
      on Release: ResetBit("Touche_Tch_Manu{90}")
      on Press: SetBit("Touche_Tch_Manu{90}")
   Button "Bouton_21" at 850,460 size 169x68; TextOff 'FERMER PORTE'
      on Release: ResetBit("Touche_Tch_Manu{91}")
      on Press: SetBit("Touche_Tch_Manu{91}")
   Rectangle "Rectangle_19" at 1034,462 size 20x20
      Appearance <- "I_porte_vision_op"
   TextField "Champ de texte_16" at 1060,460 size 137x25; Text 'Porte Ouverte'
   Rectangle "Rectangle_20" at 1034,484 size 20x20
      Appearance <- "I_porte_vision_cl"
   TextField "Champ de texte_17" at 1060,482 size 131x25; Text 'Porte Fermée'
   Rectangle "Rectangle_37" at 1034,514 size 20x20
      Appearance <- "O_Op_Porte_Vision"
   TextField "Champ de texte_32" at 1060,512 size 121x25; Text 'Ouvrir Porte'
   Rectangle "Rectangle_38" at 1034,536 size 20x20
      Appearance <- "O_Cl_porte_Vision"
   TextField "Champ de texte_33" at 1060,534 size 128x25; Text 'Fermer Porte'

screen "Mode_Manuel_Conv_carton" 1280x800, template "Modèle_Manu"
   TextField "Champ de texte_34" at 25,227 size 584x25; Text 'Convoyeur Carton - Verin de Blocage 01'
   Button "Bouton_1" at 29,268 size 169x68; TextOff 'SORTIR VERIN'
      on Release: ResetBit("Touche_Tch_Manu{80}")
      on Press: SetBit("Touche_Tch_Manu{80}")
      ObjectEnable <- "Bits_Globaux_x_Demo_Hippo_en_cours"
   Button "Bouton_3" at 210,268 size 169x68; TextOff 'RENTRER VERIN'
      on Release: ResetBit("Touche_Tch_Manu{81}")
      on Press: SetBit("Touche_Tch_Manu{81}")
      ObjectEnable <- "Bits_Globaux_x_Demo_Hippo_en_cours"
   TextField "Champ de texte_1" at 25,411 size 584x25; Text 'Convoyeur Carton - Verin de Blocage 02'
   Button "Bouton_2" at 29,452 size 169x68; TextOff 'SORTIR VERIN'
      on Release: ResetBit("Touche_Tch_Manu{82}")
      on Press: SetBit("Touche_Tch_Manu{82}")
      ObjectEnable <- "Bits_Globaux_x_Demo_Hippo_en_cours"
   Button "Bouton_4" at 210,452 size 169x68; TextOff 'RENTRER VERIN'
      on Release: ResetBit("Touche_Tch_Manu{83}")
      on Press: SetBit("Touche_Tch_Manu{83}")
      ObjectEnable <- "Bits_Globaux_x_Demo_Hippo_en_cours"
   TextField "Champ de texte_4" at 653,227 size 584x25; Text 'Convoyeur Carton - Verin de Blocage 03'
   Button "Bouton_5" at 657,268 size 169x68; TextOff 'SORTIR VERIN'
      on Release: ResetBit("Touche_Tch_Manu{84}")
      on Press: SetBit("Touche_Tch_Manu{84}")
      ObjectEnable <- "Bits_Globaux_x_Demo_Hippo_en_cours"
   Button "Bouton_6" at 838,268 size 169x68; TextOff 'RENTRER VERIN'
      on Release: ResetBit("Touche_Tch_Manu{85}")
      on Press: SetBit("Touche_Tch_Manu{85}")
      ObjectEnable <- "Bits_Globaux_x_Demo_Hippo_en_cours"
   TextField "Champ de texte_6" at 653,411 size 584x25; Text 'Convoyeur Carton - Verin de Blocage 04'
   Button "Bouton_7" at 657,452 size 169x68; TextOff 'SORTIR VERIN'
      on Release: ResetBit("Touche_Tch_Manu{86}")
      on Press: SetBit("Touche_Tch_Manu{86}")
      ObjectEnable <- "Bits_Globaux_x_Demo_Hippo_en_cours"
   Button "Bouton_8" at 838,452 size 169x68; TextOff 'RENTRER VERIN'
      on Release: ResetBit("Touche_Tch_Manu{87}")
      on Press: SetBit("Touche_Tch_Manu{87}")
      ObjectEnable <- "Bits_Globaux_x_Demo_Hippo_en_cours"
   Rectangle "Rectangle_63" at 387,270 size 20x20
      Appearance <- "I_verin_blocage_boite_sorti_01"
   TextField "Champ de texte_65" at 413,268 size 182x25; Text 'Verin bloc 01 Sorti'
   Rectangle "Rectangle_64" at 387,292 size 20x20
      Appearance <- "I_verin_blocage_boite_rentré_01"
   TextField "Champ de texte_66" at 413,290 size 199x25; Text 'Verin bloc 01 Rentré'
   Rectangle "Rectangle_65" at 390,454 size 20x20
      Appearance <- "I_verin_blocage_boite_sorti_02"
   TextField "Champ de texte_67" at 416,452 size 182x25; Text 'Verin bloc 02 Sorti'
   Rectangle "Rectangle_66" at 390,476 size 20x20
      Appearance <- "I_verin_blocage_boite_rentré_02"
   TextField "Champ de texte_68" at 416,474 size 199x25; Text 'Verin bloc 02 Rentré'
   Rectangle "Rectangle_69" at 1019,454 size 20x20
      Appearance <- "I_verin_blocage_boite_rentré_03"
   TextField "Champ de texte_71" at 1045,452 size 182x25; Text 'Verin bloc 04 Sorti'
   Rectangle "Rectangle_70" at 1019,476 size 20x20
      Appearance <- "I_verin_blocage_boite_rentré_04"
   TextField "Champ de texte_72" at 1045,474 size 199x25; Text 'Verin bloc 04 Rentré'
   Rectangle "Rectangle_2" at 1018,272 size 20x20
      Appearance <- "I_verin_blocage_boite_sorti_03"
   TextField "Champ de texte_2" at 1044,270 size 182x25; Text 'Verin bloc 03 Sorti'
   Rectangle "Rectangle_4" at 1018,294 size 20x20
      Appearance <- "I_verin_blocage_boite_sorti_04"
   TextField "Champ de texte_3" at 1044,292 size 199x25; Text 'Verin bloc 03 Rentré'
   Rectangle "Rectangle_7" at 387,330 size 20x20
      Appearance <- "O_Sortir_Blocage_boite_01"
   TextField "Champ de texte_5" at 413,328 size 114x25; Text 'Sortir Verin'
   Rectangle "Rectangle_10" at 387,352 size 20x20
      Appearance <- "O_Rentrer_Blocage_boite_01"
   TextField "Champ de texte_7" at 413,350 size 131x25; Text 'Rentrer Verin'
   Rectangle "Rectangle_11" at 390,514 size 20x20
      Appearance <- "O_Sortir_Blocage_boite_02"
   TextField "Champ de texte_8" at 416,512 size 114x25; Text 'Sortir Verin'
   Rectangle "Rectangle_12" at 390,536 size 20x20
      Appearance <- "O_Rentrer_Blocage_boite_02"
   TextField "Champ de texte_9" at 416,534 size 131x25; Text 'Rentrer Verin'
   Rectangle "Rectangle_13" at 1019,514 size 20x20
      Appearance <- "O_Sortir_Blocage_boite_04"
   TextField "Champ de texte_10" at 1045,512 size 114x25; Text 'Sortir Verin'
   Rectangle "Rectangle_14" at 1019,536 size 20x20
      Appearance <- "O_Rentrer_Blocage_boite_04"
   TextField "Champ de texte_11" at 1045,534 size 131x25; Text 'Rentrer Verin'
   Rectangle "Rectangle_15" at 1018,331 size 20x20
      Appearance <- "O_Sortir_Blocage_boite_03"
   TextField "Champ de texte_12" at 1044,329 size 114x25; Text 'Sortir Verin'
   Rectangle "Rectangle_16" at 1018,353 size 20x20
      Appearance <- "O_Rentrer_Blocage_boite_03"
   TextField "Champ de texte_13" at 1044,351 size 131x25; Text 'Rentrer Verin'

screen "Mode_Manuel_Conv_H" 1280x800, template "Modèle_Manu"
   TextField "Champ de texte_34" at 25,227 size 584x25; Text 'Hyppodrome Convoyeur 01'
   Button "Bouton_1" at 29,268 size 169x68; TextOff 'MARCHE CONVOYEUR'
      on Release: ResetBit("Touche_Tch_Manu{48}")
      on Press: SetBit("Touche_Tch_Manu{48}")
   Button "Bouton_3" at 210,268 size 169x68; TextOff 'ARRET CONVOYEUR'
      on Release: ResetBit("Touche_Tch_Manu{49}")
      on Press: SetBit("Touche_Tch_Manu{49}")
   Rectangle "Rectangle_2" at 392,279 size 20x20
      Appearance <- "I_Def_Thermique_CV01_hyppo"
   TextField "Champ de texte_2" at 418,277 size 201x25; Text 'Defaut thermique Cv'
   TextField "Champ de texte_1" at 25,411 size 584x25; Text 'Hyppodrome Convoyeur 02'
   Button "Bouton_2" at 29,452 size 169x68; TextOff 'MARCHE CONVOYEUR'
      on Release: ResetBit("Touche_Tch_Manu{50}")
      on Press: SetBit("Touche_Tch_Manu{50}")
   Button "Bouton_4" at 210,452 size 169x68; TextOff 'ARRET CONVOYEUR'
      on Release: ResetBit("Touche_Tch_Manu{51}")
      on Press: SetBit("Touche_Tch_Manu{51}")
   Rectangle "Rectangle_4" at 392,464 size 20x20
      Appearance <- "I_Def_Thermique_CV02_hyppo"
   TextField "Champ de texte_3" at 418,462 size 201x25; Text 'Defaut thermique Cv'
   TextField "Champ de texte_4" at 653,227 size 584x25; Text 'Hyppodrome Convoyeur 03'
   Button "Bouton_5" at 657,268 size 169x68; TextOff 'MARCHE CONVOYEUR'
      on Release: ResetBit("Touche_Tch_Manu{52}")
      on Press: SetBit("Touche_Tch_Manu{52}")
   Button "Bouton_6" at 838,268 size 169x68; TextOff 'ARRET CONVOYEUR'
      on Release: ResetBit("Touche_Tch_Manu{53}")
      on Press: SetBit("Touche_Tch_Manu{53}")
   Rectangle "Rectangle_7" at 1020,279 size 20x20
      Appearance <- "I_Def_Thermique_CV03_hyppo"
   TextField "Champ de texte_5" at 1046,277 size 201x25; Text 'Defaut thermique Cv'
   TextField "Champ de texte_6" at 653,411 size 584x25; Text 'Hyppodrome Convoyeur 04'
   Button "Bouton_7" at 657,452 size 169x68; TextOff 'MARCHE CONVOYEUR'
      on Release: ResetBit("Touche_Tch_Manu{54}")
      on Press: SetBit("Touche_Tch_Manu{54}")
   Button "Bouton_8" at 838,452 size 169x68; TextOff 'ARRET CONVOYEUR'
      on Release: ResetBit("Touche_Tch_Manu{55}")
      on Press: SetBit("Touche_Tch_Manu{55}")
   Rectangle "Rectangle_10" at 1020,464 size 20x20
      Appearance <- "I_Def_Thermique_CV04_hyppo"
   TextField "Champ de texte_7" at 1046,462 size 201x25; Text 'Defaut thermique Cv'
   Rectangle "Rectangle_11" at 392,304 size 20x20
      Appearance <- "Q_ON_CV_01_Hyppo"
   TextField "Champ de texte_8" at 418,302 size 180x25; Text 'Marche Convoyeur'
   Rectangle "Rectangle_12" at 392,488 size 20x20
      Appearance <- "Q_ON_CV_02_Hyppo"
   TextField "Champ de texte_9" at 418,486 size 180x25; Text 'Marche Convoyeur'
   Rectangle "Rectangle_13" at 1020,304 size 20x20
      Appearance <- "Q_ON_CV_03_Hyppo"
   TextField "Champ de texte_10" at 1047,302 size 180x25; Text 'Marche Convoyeur'
   Rectangle "Rectangle_14" at 1020,488 size 20x20
      Appearance <- "Q_ON_CV_04_Hyppo"
   TextField "Champ de texte_11" at 1046,486 size 180x25; Text 'Marche Convoyeur'
   GraphicView "Vue de graphique_3" at 240,131 size 159x86; Picture "Capture d’écran 2023-07-10 135110_1"
   Rectangle "Rectangle_15" at 260,141 size 126x11
      Appearance <- "CV01_Hipp_Marche"
   GraphicView "Vue de graphique_1" at 851,130 size 159x86; Picture "Capture d’écran 2023-07-10 135110_1"
   Rectangle "Rectangle_16" at 871,194 size 126x11
      Appearance <- "CV03_Hipp_Marche"
   GraphicView "Vue de graphique_2" at 240,580 size 159x86; Picture "Capture d’écran 2023-07-10 135110_1"
   Rectangle "Rectangle_17" at 243,588 size 18x68
      Appearance <- "CV02_Hipp_Marche"
   GraphicView "Vue de graphique_4" at 851,580 size 159x86; Picture "Capture d’écran 2023-07-10 135110_1"
   Rectangle "Rectangle_18" at 996,588 size 12x68
      Appearance <- "CV04_Hipp_Marche"

screen "Mode_Manuel_Conv_carton_01" 1280x800, template "Modèle_Manu"
   TextField "Champ de texte_34" at 44,163 size 584x25; Text 'Convoyeur Carton 01'
   Button "Bouton_1" at 48,204 size 169x68; TextOff 'MARCHE CONVOYEUR'
      on Release: ResetBit("Touche_Tch_Manu{62}")
      on Press: SetBit("Touche_Tch_Manu{62}")
   Button "Bouton_3" at 229,204 size 169x68; TextOff 'ARRET CONVOYEUR'
      on Release: ResetBit("Touche_Tch_Manu{63}")
      on Press: SetBit("Touche_Tch_Manu{63}")
   Rectangle "Rectangle_63" at 406,206 size 20x20
      Appearance <- "Var_Convoyeur_Carton_ConvoyeurC01_Marche"
   TextField "Champ de texte_65" at 432,204 size 90x25; Text 'MARCHE'
   IOField "Champ d'E/S_1" at 238,306 size 122x58; FormatPattern 9999
      ProcessValue <- "Parametres_Sp_vitesse_manu_C01"
   TextField "Champ de texte_1" at 84,317 size 160x25; Text 'VITESSE TR/MN'
   TextField "Champ de texte_2" at 85,333 size 103x25; Text '1400 Max'

screen "Mode_Manuel_Conv_carton_02" 1280x800, template "Modèle_Manu"
   TextField "Champ de texte_34" at 44,163 size 584x25; Text 'Convoyeur Carton 02'
   Button "Bouton_1" at 48,204 size 169x68; TextOff 'MARCHE CONVOYEUR'
      on Release: ResetBit("Touche_Tch_Manu{64}")
      on Press: SetBit("Touche_Tch_Manu{64}")
   Button "Bouton_3" at 229,204 size 169x68; TextOff 'ARRET CONVOYEUR'
      on Release: ResetBit("Touche_Tch_Manu{65}")
      on Press: SetBit("Touche_Tch_Manu{65}")
   Rectangle "Rectangle_63" at 406,206 size 20x20
      Appearance <- "Var_Convoyeur_Carton_ConvoyeurC02_Marche"
   TextField "Champ de texte_65" at 432,204 size 84x25; Text 'MARCHE'
   IOField "Champ d'E/S_1" at 238,306 size 122x58; FormatPattern 9999
      ProcessValue <- "Parametres_Sp_vitesse_manu_C02"
   TextField "Champ de texte_1" at 84,317 size 160x25; Text 'VITESSE TR/MN'
   TextField "Champ de texte_2" at 85,333 size 103x25; Text '1400 Max'

screen "Mode_Manuel_Conv_carton_03" 1280x800, template "Modèle_Manu"
   TextField "Champ de texte_34" at 44,163 size 584x25; Text 'Convoyeur Carton 03'
   Button "Bouton_1" at 48,204 size 169x68; TextOff 'MARCHE CONVOYEUR'
      on Release: ResetBit("Touche_Tch_Manu{66}")
      on Press: SetBit("Touche_Tch_Manu{66}")
   Button "Bouton_3" at 229,204 size 169x68; TextOff 'ARRET CONVOYEUR'
      on Release: ResetBit("Touche_Tch_Manu{67}")
      on Press: SetBit("Touche_Tch_Manu{67}")
   Rectangle "Rectangle_63" at 406,206 size 20x20
      Appearance <- "Var_Convoyeur_Carton_ConvoyeurC03_Marche"
   TextField "Champ de texte_65" at 432,204 size 84x25; Text 'MARCHE'
   IOField "Champ d'E/S_1" at 238,306 size 122x58; FormatPattern 9999
      ProcessValue <- "Parametres_Sp_vitesse_manu_C03"
   TextField "Champ de texte_1" at 84,317 size 160x25; Text 'VITESSE TR/MN'
   TextField "Champ de texte_2" at 85,333 size 103x25; Text '1400 Max'

screen "Parametrage" 1280x800, template "Modèle_1"
   Button "Bouton_3" at 1177,723 size 96x70; TextOff 'RETOUR'
      on Release: ActivateScreen("Principale", 0)
   TextField "Champ de texte_34" at 74,163 size 419x25; Text 'Convoyeur Carton 01'
   TextField "Champ de texte_1" at 95,215 size 218x25; Text 'VITESSE CONVOYEUR :'
   IOField "Champ d'E/S_1" at 303,201 size 96x51; FormatPattern 9999
      ProcessValue <- "Parametres_Sp_Vitesse_C01"
   TextField "Champ de texte_2" at 408,212 size 70x25; Text 'Tr/min'
   TextField "Champ de texte_3" at 74,287 size 419x25; Text 'Convoyeur Carton 02'
   TextField "Champ de texte_4" at 95,339 size 218x25; Text 'VITESSE CONVOYEUR :'
   IOField "Champ d'E/S_2" at 303,325 size 96x51; FormatPattern 9999
      ProcessValue <- "Parametres_Sp_Vitesse_C02"
   TextField "Champ de texte_5" at 408,336 size 70x25; Text 'Tr/min'
   TextField "Champ de texte_6" at 74,411 size 419x25; Text 'Convoyeur Carton 02'
   TextField "Champ de texte_7" at 95,463 size 218x25; Text 'VITESSE CONVOYEUR :'
   IOField "Champ d'E/S_3" at 303,449 size 96x51; FormatPattern 9999
      ProcessValue <- "Parametres_Sp_Vitesse_C03"
   TextField "Champ de texte_8" at 408,460 size 70x25; Text 'Tr/min'

screen "Visu_ES_Wieland" 1280x800, template "Modèle_ES"
   TextField "Champ de texte_1" at 43,144 size 295x25; Text 'RElAIS DE SECURITE WIELAND'
   Rectangle "Rectangle_2" at 273,244 size 20x20
      Appearance <- "I_Wieland_Au_armoire"
   TextField "Champ de texte_2" at 299,242 size 111x25; Text 'Au Armoire'
   Rectangle "Rectangle_3" at 273,266 size 20x20
      Appearance <- "I_Wieland_Au_porte01"
   TextField "Champ de texte_3" at 299,264 size 117x25; Text 'Au Porte 01'
   Rectangle "Rectangle_4" at 273,288 size 20x20
      Appearance <- "I_Wieland_Au_Porte02"
   TextField "Champ de texte_4" at 299,286 size 117x25; Text 'Au Porte 02'
   Rectangle "Rectangle_5" at 273,310 size 20x20
      Appearance <- "I_Wieland_Au_Robot01_Fanuc"
   TextField "Champ de texte_5" at 299,308 size 185x25; Text 'Au Robot 01 Fanuc'
   Rectangle "Rectangle_6" at 273,332 size 20x20
      Appearance <- "I_Wieland_Au_Robot02_Fanuc"
   TextField "Champ de texte_6" at 299,330 size 185x25; Text 'Au Robot 02 Fanuc'
   Rectangle "Rectangle_7" at 273,354 size 20x20
      Appearance <- "I_Wieland_Au_Robot03_ABB"
   TextField "Champ de texte_7" at 299,352 size 168x25; Text 'Au Robot 03 ABB'
   Rectangle "Rectangle_8" at 273,376 size 20x20
      Appearance <- "I_Wielmand_Au_Robot04_UR"
   TextField "Champ de texte_8" at 299,374 size 156x25; Text 'Au Robot 04 UR'
   Rectangle "Rectangle_9" at 273,398 size 20x20
      Appearance <- "I_Wieland_Au_Robot05_UR"
   TextField "Champ de texte_9" at 299,396 size 156x25; Text 'Au Robot 05 UR'
   Rectangle "Rectangle_10" at 483,244 size 20x20
      Appearance <- "I_wieland_Au_Carroussel"
   TextField "Champ de texte_10" at 509,242 size 157x25; Text 'Au Hyppodrome'
   Rectangle "Rectangle_11" at 483,266 size 20x20
      Appearance <- "I_Wieland_Au_Carterisation"
   TextField "Champ de texte_11" at 509,264 size 165x25; Text 'Au Carterisation'
   Rectangle "Rectangle_12" at 483,288 size 20x20
      Appearance <- "I_Wieland_Porte 01 ouverte"
   TextField "Champ de texte_12" at 509,286 size 158x25; Text 'Porte 01 fermée'
   Rectangle "Rectangle_13" at 483,310 size 20x20
      Appearance <- "I_Wieland_Porte 02 Ouverte"
   TextField "Champ de texte_13" at 509,308 size 158x25; Text 'Porte 02 fermée'
   Rectangle "Rectangle_14" at 483,332 size 20x20
      Appearance <- "I_Wieland_Rearmement"
   TextField "Champ de texte_14" at 509,330 size 124x25; Text 'Rearmement'
   Rectangle "Rectangle_15" at 483,354 size 20x20
      Appearance <- "I_Wieland_Dmd acces"
   TextField "Champ de texte_15" at 509,352 size 151x25; Text 'Demande acces'
   Rectangle "Rectangle_16" at 483,376 size 20x20
      Appearance <- "I_Wieland_Mise sous puissance"
   TextField "Champ de texte_16" at 509,374 size 198x25; Text 'Mise sous puissance'
   Rectangle "Rectangle_17" at 483,398 size 20x20
      Appearance <- "I_Wieland_Mise hors puissance"
   TextField "Champ de texte_17" at 509,396 size 196x25; Text 'Mise hors puissance'
   TextField "Champ de texte_34" at 254,173 size 880x25; Text 'ENTREES PLC --- SORTIES WIELAND'
   TextField "Champ de texte_35" at 273,219 size 59x25; Text '%I16'
   TextField "Champ de texte_37" at 483,219 size 59x25; Text '%I17'
   Rectangle "Rectangle_18" at 692,244 size 20x20
      Appearance <- "I_Wieland_Acces_autorisé"
   TextField "Champ de texte_18" at 718,242 size 145x25; Text 'Acces Autorisé'
   Rectangle "Rectangle_19" at 692,266 size 20x20
      Appearance <- "I_Wieland_rearmement_Porte"
   TextField "Champ de texte_19" at 718,264 size 181x25; Text 'Rearmement Porte'
   Rectangle "Rectangle_20" at 692,288 size 20x20
      Appearance <- "I_Wieland_En_Service"
   TextField "Champ de texte_20" at 718,286 size 103x25; Text 'En Service'
   Rectangle "Rectangle_21" at 692,310 size 20x20
      Appearance <- "I_Wieland_Porte_non_Réarmée"
   TextField "Champ de texte_21" at 718,308 size 186x25; Text 'Porte non Rearmée'
   Rectangle "Rectangle_22" at 692,332 size 20x20
      Appearance <- "AlwaysFALSE"
   TextField "Champ de texte_22" at 718,330 size 53x25; Text 'Libre'
   Rectangle "Rectangle_23" at 692,354 size 20x20
      Appearance <- "AlwaysFALSE"
   TextField "Champ de texte_23" at 718,352 size 53x25; Text 'Libre'
   Rectangle "Rectangle_24" at 692,376 size 20x20
      Appearance <- "AlwaysFALSE"
   TextField "Champ de texte_24" at 718,374 size 53x25; Text 'Libre'
   Rectangle "Rectangle_25" at 692,398 size 20x20
      Appearance <- "AlwaysFALSE"
   TextField "Champ de texte_25" at 718,396 size 53x25; Text 'Libre'
   Rectangle "Rectangle_26" at 902,244 size 20x20
      Appearance <- "AlwaysFALSE"
   TextField "Champ de texte_26" at 928,242 size 53x25; Text 'Libre'
   Rectangle "Rectangle_27" at 902,266 size 20x20
      Appearance <- "AlwaysFALSE"
   TextField "Champ de texte_27" at 928,264 size 53x25; Text 'Libre'
   Rectangle "Rectangle_28" at 902,288 size 20x20
      Appearance <- "AlwaysFALSE"
   TextField "Champ de texte_28" at 928,286 size 53x25; Text 'Libre'
   Rectangle "Rectangle_29" at 902,310 size 20x20
      Appearance <- "AlwaysFALSE"
   TextField "Champ de texte_29" at 928,308 size 53x25; Text 'Libre'
   Rectangle "Rectangle_30" at 902,332 size 20x20
      Appearance <- "AlwaysFALSE"
   TextField "Champ de texte_30" at 928,330 size 53x25; Text 'Libre'
   Rectangle "Rectangle_31" at 902,354 size 20x20
      Appearance <- "AlwaysFALSE"
   TextField "Champ de texte_31" at 928,352 size 53x25; Text 'Libre'
   Rectangle "Rectangle_32" at 902,376 size 20x20
      Appearance <- "AlwaysFALSE"
   TextField "Champ de texte_32" at 928,374 size 53x25; Text 'Libre'
   Rectangle "Rectangle_34" at 902,398 size 20x20
      Appearance <- "AlwaysFALSE"
   TextField "Champ de texte_33" at 928,396 size 53x25; Text 'Libre'
   TextField "Champ de texte_36" at 692,219 size 59x25; Text '%I18'
   TextField "Champ de texte_38" at 902,219 size 59x25; Text '%I19'
   GraphicView "Vue de graphique_1" at 65,187 size 147x117; Picture "Sans titre"
   Rectangle "Rectangle_37" at 273,519 size 20x20
      Appearance <- "Q_Wieland_Acces_Autorisé"
   TextField "Champ de texte_39" at 299,517 size 202x25; Text 'Acces Porte Autorisé'
   Rectangle "Rectangle_38" at 273,541 size 20x20
      Appearance <- "AlwaysFALSE"
   TextField "Champ de texte_40" at 299,539 size 53x25; Text 'Libre'
   Rectangle "Rectangle_39" at 273,563 size 20x20
      Appearance <- "AlwaysFALSE"
   TextField "Champ de texte_41" at 299,561 size 53x25; Text 'Libre'
   Rectangle "Rectangle_40" at 273,585 size 20x20
      Appearance <- "AlwaysFALSE"
   TextField "Champ de texte_42" at 299,583 size 53x25; Text 'Libre'
   Rectangle "Rectangle_41" at 273,607 size 20x20
      Appearance <- "AlwaysFALSE"
   TextField "Champ de texte_43" at 299,605 size 53x25; Text 'Libre'
   Rectangle "Rectangle_42" at 273,629 size 20x20
      Appearance <- "AlwaysFALSE"
   TextField "Champ de texte_44" at 299,627 size 53x25; Text 'Libre'
   Rectangle "Rectangle_43" at 273,651 size 20x20
      Appearance <- "AlwaysFALSE"
   TextField "Champ de texte_45" at 299,649 size 53x25; Text 'Libre'
   Rectangle "Rectangle_44" at 273,673 size 20x20
      Appearance <- "AlwaysFALSE"
   TextField "Champ de texte_46" at 299,671 size 53x25; Text 'Libre'
   Rectangle "Rectangle_45" at 483,519 size 20x20
      Appearance <- "AlwaysFALSE"
   TextField "Champ de texte_47" at 509,517 size 53x25; Text 'Libre'
   Rectangle "Rectangle_46" at 483,541 size 20x20
      Appearance <- "AlwaysFALSE"
   TextField "Champ de texte_48" at 509,539 size 53x25; Text 'Libre'
   Rectangle "Rectangle_47" at 483,563 size 20x20
      Appearance <- "AlwaysFALSE"
   TextField "Champ de texte_49" at 509,561 size 53x25; Text 'Libre'
   Rectangle "Rectangle_48" at 483,585 size 20x20
      Appearance <- "AlwaysFALSE"
   TextField "Champ de texte_50" at 509,583 size 53x25; Text 'Libre'
   Rectangle "Rectangle_49" at 483,607 size 20x20
      Appearance <- "AlwaysFALSE"
   TextField "Champ de texte_51" at 509,605 size 53x25; Text 'Libre'
   Rectangle "Rectangle_50" at 483,629 size 20x20
      Appearance <- "AlwaysFALSE"
   TextField "Champ de texte_52" at 509,627 size 53x25; Text 'Libre'
   Rectangle "Rectangle_51" at 483,651 size 20x20
      Appearance <- "AlwaysFALSE"
   TextField "Champ de texte_53" at 509,649 size 53x25; Text 'Libre'
   Rectangle "Rectangle_52" at 483,673 size 20x20
      Appearance <- "AlwaysFALSE"
   TextField "Champ de texte_54" at 509,671 size 53x25; Text 'Libre'
   TextField "Champ de texte_55" at 254,448 size 880x25; Text 'SORTIES PLC --- ENTREES WIELAND'
   TextField "Champ de texte_56" at 273,494 size 64x25; Text '%Q18'
   TextField "Champ de texte_57" at 483,494 size 64x25; Text '%Q19'
   Rectangle "Rectangle_54" at 692,519 size 20x20
      Appearance <- "AlwaysFALSE"
   TextField "Champ de texte_58" at 718,517 size 53x25; Text 'Libre'
   Rectangle "Rectangle_55" at 692,541 size 20x20
      Appearance <- "AlwaysFALSE"
   TextField "Champ de texte_59" at 718,539 size 53x25; Text 'Libre'
   Rectangle "Rectangle_56" at 692,563 size 20x20
      Appearance <- "AlwaysFALSE"
   TextField "Champ de texte_60" at 718,561 size 53x25; Text 'Libre'
   Rectangle "Rectangle_57" at 692,585 size 20x20
      Appearance <- "AlwaysFALSE"
   TextField "Champ de texte_61" at 718,583 size 53x25; Text 'Libre'
   Rectangle "Rectangle_58" at 692,607 size 20x20
      Appearance <- "AlwaysFALSE"
   TextField "Champ de texte_62" at 718,605 size 53x25; Text 'Libre'
   Rectangle "Rectangle_59" at 692,629 size 20x20
      Appearance <- "AlwaysFALSE"
   TextField "Champ de texte_63" at 718,627 size 53x25; Text 'Libre'
   Rectangle "Rectangle_60" at 692,651 size 20x20
      Appearance <- "AlwaysFALSE"
   TextField "Champ de texte_64" at 718,649 size 53x25; Text 'Libre'
   Rectangle "Rectangle_61" at 692,673 size 20x20
      Appearance <- "AlwaysFALSE"
   TextField "Champ de texte_65" at 718,671 size 53x25; Text 'Libre'
   Rectangle "Rectangle_62" at 902,519 size 20x20
      Appearance <- "AlwaysFALSE"
   TextField "Champ de texte_66" at 928,517 size 53x25; Text 'Libre'
   Rectangle "Rectangle_63" at 902,541 size 20x20
      Appearance <- "AlwaysFALSE"
   TextField "Champ de texte_67" at 928,539 size 53x25; Text 'Libre'
   Rectangle "Rectangle_64" at 902,563 size 20x20
      Appearance <- "AlwaysFALSE"
   TextField "Champ de texte_68" at 928,561 size 53x25; Text 'Libre'
   Rectangle "Rectangle_65" at 902,585 size 20x20
      Appearance <- "AlwaysFALSE"
   TextField "Champ de texte_69" at 928,583 size 53x25; Text 'Libre'
   Rectangle "Rectangle_66" at 902,607 size 20x20
      Appearance <- "AlwaysFALSE"
   TextField "Champ de texte_70" at 928,605 size 53x25; Text 'Libre'
   Rectangle "Rectangle_67" at 902,629 size 20x20
      Appearance <- "AlwaysFALSE"
   TextField "Champ de texte_71" at 928,627 size 53x25; Text 'Libre'
   Rectangle "Rectangle_68" at 902,651 size 20x20
      Appearance <- "AlwaysFALSE"
   TextField "Champ de texte_72" at 928,649 size 53x25; Text 'Libre'
   Rectangle "Rectangle_69" at 902,673 size 20x20
      Appearance <- "AlwaysFALSE"
   TextField "Champ de texte_73" at 928,671 size 53x25; Text 'Libre'
   TextField "Champ de texte_74" at 692,494 size 64x25; Text '%Q20'
   TextField "Champ de texte_75" at 902,494 size 64x25; Text '%Q21'

screen "Visu_ES_Variateur_C1" 1280x800, template "Modèle_ES"
   Rectangle "Rectangle_2" at 204,218 size 20x20
      Appearance <- "Var_Convoyeur_Carton_ConvoyeurC01_Reserve01"
   TextField "Champ de texte_2" at 230,216 size 110x25; Text 'Reserve 01'
   Rectangle "Rectangle_3" at 204,240 size 20x20
      Appearance <- "Var_Convoyeur_Carton_ConvoyeurC01_Reserve02"
   TextField "Champ de texte_3" at 230,238 size 110x25; Text 'Reserve 02'
   Rectangle "Rectangle_4" at 204,262 size 20x20
      Appearance <- "Var_Convoyeur_Carton_ConvoyeurC01_PilotageParApi"
   TextField "Champ de texte_4" at 230,260 size 120x25; Text 'Pilotage Api'
   Rectangle "Rectangle_5" at 204,284 size 20x20
      Appearance <- "Var_Convoyeur_Carton_ConvoyeurC01_InversionConsigne"
   TextField "Champ de texte_5" at 230,282 size 189x25; Text 'Inversion Consigne'
   Rectangle "Rectangle_6" at 204,306 size 20x20
      Appearance <- "Var_Convoyeur_Carton_ConvoyeurC01_Reserve03"
   TextField "Champ de texte_6" at 230,304 size 110x25; Text 'Reserve 03'
   Rectangle "Rectangle_7" at 204,328 size 20x20
      Appearance <- "Var_Convoyeur_Carton_ConvoyeurC01_PotPlus"
   TextField "Champ de texte_7" at 230,326 size 83x25; Text 'Pot Plus'
   Rectangle "Rectangle_8" at 204,350 size 20x20
      Appearance <- "Var_Convoyeur_Carton_ConvoyeurC01_PotMoins"
   TextField "Champ de texte_8" at 230,348 size 99x25; Text 'Pot Moins'
   Rectangle "Rectangle_9" at 204,372 size 20x20
      Appearance <- "Var_Convoyeur_Carton_ConvoyeurC01_Reserve04"
   TextField "Champ de texte_9" at 230,370 size 110x25; Text 'Reserve 04'
   TextField "Champ de texte_34" at 185,147 size 347x25; Text 'ENTREES'
   TextField "Champ de texte_35" at 204,193 size 90x25; Text '%QD256'
   GraphicView "Vue de graphique_1" at 39,160 size 112x173; Picture "Graphique_6"
   Rectangle "Rectangle_36" at 204,395 size 20x20
      Appearance <- "Var_Convoyeur_Carton_ConvoyeurC01_Marche"
   TextField "Champ de texte_1" at 230,393 size 73x25; Text 'Marche'
   Rectangle "Rectangle_37" at 204,417 size 20x20
      Appearance <- "Var_Convoyeur_Carton_ConvoyeurC01_Arret2"
   TextField "Champ de texte_39" at 230,415 size 71x25; Text 'Arret 2'
   Rectangle "Rectangle_38" at 204,439 size 20x20
      Appearance <- "Var_Convoyeur_Carton_ConvoyeurC01_Arret3"
   TextField "Champ de texte_40" at 230,437 size 71x25; Text 'Arret 3'
   Rectangle "Rectangle_39" at 204,461 size 20x20
      Appearance <- "Var_Convoyeur_Carton_ConvoyeurC01_DebloqFonctionnement"
   Rectangle "Rectangle_40" at 204,483 size 20x20
      Appearance <- "Var_Convoyeur_Carton_ConvoyeurC01_DebloqRampe"
   TextField "Champ de texte_41" at 230,481 size 142x25; Text 'Debloq Rampe'
   Rectangle "Rectangle_41" at 204,505 size 20x20
      Appearance <- "Var_Convoyeur_Carton_ConvoyeurC01_GelerGenerateurRampe"
   TextField "Champ de texte_42" at 230,503 size 179x25; Text 'Geler Gene Rampe'
   Rectangle "Rectangle_42" at 204,527 size 20x20
      Appearance <- "Var_Convoyeur_Carton_ConvoyeurC01_DebloqConsigne"
   TextField "Champ de texte_43" at 230,525 size 165x25; Text 'Debloq Consigne'
   Rectangle "Rectangle_43" at 204,549 size 20x20
      Appearance <- "Var_Convoyeur_Carton_ConvoyeurC01_AcquitDefaut"
   TextField "Champ de texte_44" at 230,547 size 134x25; Text 'Acquit defaut'
   TextField "Champ de texte_45" at 230,461 size 158x25; Text 'Debloq fonction'
   IOField "Champ d'E/S_1" at 212,607 size 109x32; FormatPattern s99999
      ProcessValue <- "Var_Convoyeur_Carton_ConvoyeurC01_Consigne"
   TextField "Champ de texte_46" at 216,582 size 92x25; Text 'Consigne'
   Rectangle "Rectangle_11" at 590,217 size 20x20
      Appearance <- "Var_Convoyeur_Carton_ConvoyeurC01_EcartVitesse"
   TextField "Champ de texte_10" at 616,215 size 127x25; Text 'Ecart Vitesse'
   Rectangle "Rectangle_12" at 590,239 size 20x20
      Appearance <- "Var_Convoyeur_Carton_ConvoyeurC01_CommandeDemander"
   TextField "Champ de texte_11" at 616,237 size 212x25; Text 'Commande demandée'
   Rectangle "Rectangle_13" at 590,261 size 20x20
      Appearance <- "Var_Convoyeur_Carton_ConvoyeurC01_VitesseMaxAtteinte"
   TextField "Champ de texte_12" at 616,259 size 199x25; Text 'Vitesse max atteinte'
   Rectangle "Rectangle_14" at 590,283 size 20x20
      Appearance <- "Var_Convoyeur_Carton_ConvoyeurC01_Limite"
   TextField "Champ de texte_13" at 616,281 size 182x25; Text 'Limites de courant'
   Rectangle "Rectangle_15" at 590,305 size 20x20
      Appearance <- "Var_Convoyeur_Carton_ConvoyeurC01_FreinMoteur"
   TextField "Champ de texte_14" at 616,303 size 126x25; Text 'Frein Moteur'
   Rectangle "Rectangle_16" at 590,327 size 20x20
      Appearance <- "Var_Convoyeur_Carton_ConvoyeurC01_AlarmeSurchauffe"
   TextField "Champ de texte_15" at 616,325 size 181x25; Text 'Alarme Surchauffe'
   Rectangle "Rectangle_17" at 590,349 size 20x20
      Appearance <- "Var_Convoyeur_Carton_ConvoyeurC01_MoteurSensAvant"
   TextField "Champ de texte_16" at 616,347 size 180x25; Text 'Moteur sens avant'
   Rectangle "Rectangle_18" at 590,371 size 20x20
      Appearance <- "Var_Convoyeur_Carton_ConvoyeurC01_SurchargeMoteur"
   TextField "Champ de texte_17" at 616,369 size 174x25; Text 'Surcharge Moteur'
   TextField "Champ de texte_18" at 571,146 size 347x25; Text 'SORTIES'
   TextField "Champ de texte_19" at 590,192 size 85x25; Text '%ID256'
   Rectangle "Rectangle_20" at 590,394 size 20x20
      Appearance <- "Var_Convoyeur_Carton_ConvoyeurC01_PretEnclenchement"
   TextField "Champ de texte_20" at 616,392 size 193x25; Text 'Pret enclenchement'
   Rectangle "Rectangle_21" at 590,416 size 20x20
      Appearance <- "Var_Convoyeur_Carton_ConvoyeurC01_PretFonctionnement"
   TextField "Champ de texte_21" at 616,414 size 210x25; Text 'Pret Fonctionnement'
   Rectangle "Rectangle_22" at 590,438 size 20x20
      Appearance <- "Var_Convoyeur_Carton_ConvoyeurC01_Fonctionnement_Debloq"
   TextField "Champ de texte_22" at 616,436 size 236x25; Text 'Fonctionnement debloq.'
   Rectangle "Rectangle_23" at 590,460 size 20x20
      Appearance <- "Var_Convoyeur_Carton_ConvoyeurC01_DefautActif"
   Rectangle "Rectangle_24" at 590,482 size 20x20
      Appearance <- "Var_Convoyeur_Carton_ConvoyeurC01_Arret2Etat"
   TextField "Champ de texte_23" at 616,480 size 138x25; Text 'Arret 2 inactif'
   Rectangle "Rectangle_25" at 590,504 size 20x20
      Appearance <- "Var_Convoyeur_Carton_ConvoyeurC01_Arret3Etat"
   TextField "Champ de texte_24" at 616,502 size 138x25; Text 'Arret 3 inactif'
   Rectangle "Rectangle_26" at 590,526 size 20x20
      Appearance <- "Var_Convoyeur_Carton_ConvoyeurC01_BlocageActif"
   TextField "Champ de texte_25" at 616,524 size 135x25; Text 'Blocage actif'
   Rectangle "Rectangle_27" at 590,548 size 20x20
      Appearance <- "Var_Convoyeur_Carton_ConvoyeurC01_AlarmeActive"
   TextField "Champ de texte_26" at 616,546 size 134x25; Text 'Alarme active'
   TextField "Champ de texte_27" at 616,460 size 118x25; Text 'Défaut actif'
   IOField "Champ d'E/S_2" at 598,606 size 96x32; FormatPattern s99999
      ProcessValue <- "Var_Convoyeur_Carton_ConvoyeurC01_Vitesse"
   TextField "Champ de texte_28" at 602,581 size 73x25; Text 'Vitesse'
   Button "Bouton_1" at 8,8 size 96x32; TextOff 'Text'
   Button "Bouton_2" at 26,386 size 140x53; TextOff 'Convoyeur 01'
      on Release: ActivateScreen("Visu_ES_Variateur_C1", 0)
   Button "Bouton_3" at 25,450 size 140x53; TextOff 'Convoyeur 02'
      on Release: ActivateScreen("Visu_ES_Variateur_C2", 0)
   Button "Bouton_4" at 25,514 size 140x53; TextOff 'Convoyeur 03'
      on Release: ActivateScreen("Visu_ES_Variateur_C3", 0)

screen "Visu_ES_Variateur_C2" 1280x800, template "Modèle_ES"
   Rectangle "Rectangle_2" at 204,218 size 20x20
      Appearance <- "Var_Convoyeur_Carton_ConvoyeurC02_Reserve01"
   TextField "Champ de texte_2" at 230,216 size 110x25; Text 'Reserve 01'
   Rectangle "Rectangle_3" at 204,240 size 20x20
      Appearance <- "Var_Convoyeur_Carton_ConvoyeurC02_Reserve02"
   TextField "Champ de texte_3" at 230,238 size 110x25; Text 'Reserve 02'
   Rectangle "Rectangle_4" at 204,262 size 20x20
      Appearance <- "Var_Convoyeur_Carton_ConvoyeurC02_PilotageParApi"
   TextField "Champ de texte_4" at 230,260 size 120x25; Text 'Pilotage Api'
   Rectangle "Rectangle_5" at 204,284 size 20x20
      Appearance <- "Var_Convoyeur_Carton_ConvoyeurC02_InversionConsigne"
   TextField "Champ de texte_5" at 230,282 size 189x25; Text 'Inversion Consigne'
   Rectangle "Rectangle_6" at 204,306 size 20x20
      Appearance <- "Var_Convoyeur_Carton_ConvoyeurC02_Reserve03"
   TextField "Champ de texte_6" at 230,304 size 110x25; Text 'Reserve 03'
   Rectangle "Rectangle_7" at 204,328 size 20x20
      Appearance <- "Var_Convoyeur_Carton_ConvoyeurC02_PotPlus"
   TextField "Champ de texte_7" at 230,326 size 83x25; Text 'Pot Plus'
   Rectangle "Rectangle_8" at 204,350 size 20x20
      Appearance <- "Var_Convoyeur_Carton_ConvoyeurC02_PotMoins"
   TextField "Champ de texte_8" at 230,348 size 99x25; Text 'Pot Moins'
   Rectangle "Rectangle_9" at 204,372 size 20x20
      Appearance <- "Var_Convoyeur_Carton_ConvoyeurC02_Reserve04"
   TextField "Champ de texte_9" at 230,370 size 110x25; Text 'Reserve 04'
   TextField "Champ de texte_34" at 185,147 size 347x25; Text 'ENTREES'
   TextField "Champ de texte_35" at 204,193 size 90x25; Text '%QD260'
   GraphicView "Vue de graphique_1" at 39,160 size 112x173; Picture "Graphique_6"
   Rectangle "Rectangle_36" at 204,395 size 20x20
      Appearance <- "Var_Convoyeur_Carton_ConvoyeurC02_Marche"
   TextField "Champ de texte_1" at 230,393 size 73x25; Text 'Marche'
   Rectangle "Rectangle_37" at 204,417 size 20x20
      Appearance <- "Var_Convoyeur_Carton_ConvoyeurC02_Arret2"
   TextField "Champ de texte_39" at 230,415 size 71x25; Text 'Arret 2'
   Rectangle "Rectangle_38" at 204,439 size 20x20
      Appearance <- "Var_Convoyeur_Carton_ConvoyeurC02_Arret3"
   TextField "Champ de texte_40" at 230,437 size 71x25; Text 'Arret 3'
   Rectangle "Rectangle_39" at 204,461 size 20x20
      Appearance <- "Var_Convoyeur_Carton_ConvoyeurC02_DebloqFonctionnement"
   Rectangle "Rectangle_40" at 204,483 size 20x20
      Appearance <- "Var_Convoyeur_Carton_ConvoyeurC02_DebloqRampe"
   TextField "Champ de texte_41" at 230,481 size 142x25; Text 'Debloq Rampe'
   Rectangle "Rectangle_41" at 204,505 size 20x20
      Appearance <- "Var_Convoyeur_Carton_ConvoyeurC02_GelerGenerateurRampe"
   TextField "Champ de texte_42" at 230,503 size 179x25; Text 'Geler Gene Rampe'
   Rectangle "Rectangle_42" at 204,527 size 20x20
      Appearance <- "Var_Convoyeur_Carton_ConvoyeurC02_DebloqConsigne"
   TextField "Champ de texte_43" at 230,525 size 165x25; Text 'Debloq Consigne'
   Rectangle "Rectangle_43" at 204,549 size 20x20
      Appearance <- "Var_Convoyeur_Carton_ConvoyeurC02_AcquitDefaut"
   TextField "Champ de texte_44" at 230,547 size 134x25; Text 'Acquit defaut'
   TextField "Champ de texte_45" at 230,461 size 158x25; Text 'Debloq fonction'
   IOField "Champ d'E/S_1" at 212,607 size 109x32; FormatPattern s99999
      ProcessValue <- "Var_Convoyeur_Carton_ConvoyeurC02_Consigne"
   TextField "Champ de texte_46" at 216,582 size 92x25; Text 'Consigne'
   Rectangle "Rectangle_11" at 590,217 size 20x20
      Appearance <- "Var_Convoyeur_Carton_ConvoyeurC02_EcartVitesse"
   TextField "Champ de texte_10" at 616,215 size 127x25; Text 'Ecart Vitesse'
   Rectangle "Rectangle_12" at 590,239 size 20x20
      Appearance <- "Var_Convoyeur_Carton_ConvoyeurC02_CommandeDemander"
   TextField "Champ de texte_11" at 616,237 size 212x25; Text 'Commande demandée'
   Rectangle "Rectangle_13" at 590,261 size 20x20
      Appearance <- "Var_Convoyeur_Carton_ConvoyeurC02_VitesseMaxAtteinte"
   TextField "Champ de texte_12" at 616,259 size 199x25; Text 'Vitesse max atteinte'
   Rectangle "Rectangle_14" at 590,283 size 20x20
      Appearance <- "Var_Convoyeur_Carton_ConvoyeurC02_Limite"
   TextField "Champ de texte_13" at 616,281 size 182x25; Text 'Limites de courant'
   Rectangle "Rectangle_15" at 590,305 size 20x20
      Appearance <- "Var_Convoyeur_Carton_ConvoyeurC02_FreinMoteur"
   TextField "Champ de texte_14" at 616,303 size 126x25; Text 'Frein Moteur'
   Rectangle "Rectangle_16" at 590,327 size 20x20
      Appearance <- "Var_Convoyeur_Carton_ConvoyeurC02_AlarmeSurchauffe"
   TextField "Champ de texte_15" at 616,325 size 181x25; Text 'Alarme Surchauffe'
   Rectangle "Rectangle_17" at 590,349 size 20x20
      Appearance <- "Var_Convoyeur_Carton_ConvoyeurC02_MoteurSensAvant"
   TextField "Champ de texte_16" at 616,347 size 180x25; Text 'Moteur sens avant'
   Rectangle "Rectangle_18" at 590,371 size 20x20
      Appearance <- "Var_Convoyeur_Carton_ConvoyeurC02_SurchargeMoteur"
   TextField "Champ de texte_17" at 616,369 size 174x25; Text 'Surcharge Moteur'
   TextField "Champ de texte_18" at 571,146 size 347x25; Text 'SORTIES'
   TextField "Champ de texte_19" at 590,192 size 85x25; Text '%ID260'
   Rectangle "Rectangle_20" at 590,394 size 20x20
      Appearance <- "Var_Convoyeur_Carton_ConvoyeurC02_PretEnclenchement"
   TextField "Champ de texte_20" at 616,392 size 193x25; Text 'Pret enclenchement'
   Rectangle "Rectangle_21" at 590,416 size 20x20
      Appearance <- "Var_Convoyeur_Carton_ConvoyeurC02_PretFonctionnement"
   TextField "Champ de texte_21" at 616,414 size 210x25; Text 'Pret Fonctionnement'
   Rectangle "Rectangle_22" at 590,438 size 20x20
      Appearance <- "Var_Convoyeur_Carton_ConvoyeurC02_Fonctionnement_Debloq"
   TextField "Champ de texte_22" at 616,436 size 236x25; Text 'Fonctionnement debloq.'
   Rectangle "Rectangle_23" at 590,460 size 20x20
      Appearance <- "Var_Convoyeur_Carton_ConvoyeurC02_DefautActif"
   Rectangle "Rectangle_24" at 590,482 size 20x20
      Appearance <- "Var_Convoyeur_Carton_ConvoyeurC02_Arret2Etat"
   TextField "Champ de texte_23" at 616,480 size 138x25; Text 'Arret 2 inactif'
   Rectangle "Rectangle_25" at 590,504 size 20x20
      Appearance <- "Var_Convoyeur_Carton_ConvoyeurC02_Arret3Etat"
   TextField "Champ de texte_24" at 616,502 size 138x25; Text 'Arret 3 inactif'
   Rectangle "Rectangle_26" at 590,526 size 20x20
      Appearance <- "Var_Convoyeur_Carton_ConvoyeurC02_BlocageActif"
   TextField "Champ de texte_25" at 616,524 size 135x25; Text 'Blocage actif'
   Rectangle "Rectangle_27" at 590,548 size 20x20
      Appearance <- "Var_Convoyeur_Carton_ConvoyeurC02_AlarmeActive"
   TextField "Champ de texte_26" at 616,546 size 134x25; Text 'Alarme active'
   TextField "Champ de texte_27" at 616,460 size 118x25; Text 'Défaut actif'
   IOField "Champ d'E/S_2" at 598,606 size 96x32; FormatPattern s99999
      ProcessValue <- "Var_Convoyeur_Carton_ConvoyeurC02_Vitesse"
   TextField "Champ de texte_28" at 602,581 size 73x25; Text 'Vitesse'
   Button "Bouton_1" at 8,8 size 96x32; TextOff 'Text'
   Button "Bouton_2" at 26,386 size 140x53; TextOff 'Convoyeur 01'
      on Release: ActivateScreen("Visu_ES_Variateur_C1", 0)
   Button "Bouton_3" at 25,450 size 140x53; TextOff 'Convoyeur 02'
      on Release: ActivateScreen("Visu_ES_Variateur_C2", 0)
   Button "Bouton_4" at 25,514 size 140x53; TextOff 'Convoyeur 03'
      on Release: ActivateScreen("Visu_ES_Variateur_C3", 0)

screen "Visu_ES_Variateur_C3" 1280x800, template "Modèle_ES"
   Rectangle "Rectangle_2" at 204,218 size 20x20
      Appearance <- "Var_Convoyeur_Carton_ConvoyeurC03_Reserve01"
   TextField "Champ de texte_2" at 230,216 size 110x25; Text 'Reserve 01'
   Rectangle "Rectangle_3" at 204,240 size 20x20
      Appearance <- "Var_Convoyeur_Carton_ConvoyeurC03_Reserve02"
   TextField "Champ de texte_3" at 230,238 size 110x25; Text 'Reserve 02'
   Rectangle "Rectangle_4" at 204,262 size 20x20
      Appearance <- "Var_Convoyeur_Carton_ConvoyeurC03_PilotageParApi"
   TextField "Champ de texte_4" at 230,260 size 120x25; Text 'Pilotage Api'
   Rectangle "Rectangle_5" at 204,284 size 20x20
      Appearance <- "Var_Convoyeur_Carton_ConvoyeurC03_InversionConsigne"
   TextField "Champ de texte_5" at 230,282 size 189x25; Text 'Inversion Consigne'
   Rectangle "Rectangle_6" at 204,306 size 20x20
      Appearance <- "Var_Convoyeur_Carton_ConvoyeurC03_Reserve03"
   TextField "Champ de texte_6" at 230,304 size 110x25; Text 'Reserve 03'
   Rectangle "Rectangle_7" at 204,328 size 20x20
      Appearance <- "Var_Convoyeur_Carton_ConvoyeurC03_PotPlus"
   TextField "Champ de texte_7" at 230,326 size 83x25; Text 'Pot Plus'
   Rectangle "Rectangle_8" at 204,350 size 20x20
      Appearance <- "Var_Convoyeur_Carton_ConvoyeurC03_PotMoins"
   TextField "Champ de texte_8" at 230,348 size 99x25; Text 'Pot Moins'
   Rectangle "Rectangle_9" at 204,372 size 20x20
      Appearance <- "Var_Convoyeur_Carton_ConvoyeurC03_Reserve04"
   TextField "Champ de texte_9" at 230,370 size 110x25; Text 'Reserve 04'
   TextField "Champ de texte_34" at 185,147 size 347x25; Text 'ENTREES'
   TextField "Champ de texte_35" at 204,193 size 90x25; Text '%QD264'
   GraphicView "Vue de graphique_1" at 39,160 size 112x173; Picture "Graphique_6"
   Rectangle "Rectangle_36" at 204,395 size 20x20
      Appearance <- "Var_Convoyeur_Carton_ConvoyeurC03_Marche"
   TextField "Champ de texte_1" at 230,393 size 73x25; Text 'Marche'
   Rectangle "Rectangle_37" at 204,417 size 20x20
      Appearance <- "Var_Convoyeur_Carton_ConvoyeurC03_Arret2"
   TextField "Champ de texte_39" at 230,415 size 71x25; Text 'Arret 2'
   Rectangle "Rectangle_38" at 204,439 size 20x20
      Appearance <- "Var_Convoyeur_Carton_ConvoyeurC03_Arret3"
   TextField "Champ de texte_40" at 230,437 size 71x25; Text 'Arret 3'
   Rectangle "Rectangle_39" at 204,461 size 20x20
      Appearance <- "Var_Convoyeur_Carton_ConvoyeurC03_DebloqFonctionnement"
   Rectangle "Rectangle_40" at 204,483 size 20x20
      Appearance <- "Var_Convoyeur_Carton_ConvoyeurC03_DebloqRampe"
   TextField "Champ de texte_41" at 230,481 size 142x25; Text 'Debloq Rampe'
   Rectangle "Rectangle_41" at 204,505 size 20x20
      Appearance <- "Var_Convoyeur_Carton_ConvoyeurC03_GelerGenerateurRampe"
   TextField "Champ de texte_42" at 230,503 size 179x25; Text 'Geler Gene Rampe'
   Rectangle "Rectangle_42" at 204,527 size 20x20
      Appearance <- "Var_Convoyeur_Carton_ConvoyeurC03_DebloqConsigne"
   TextField "Champ de texte_43" at 230,525 size 165x25; Text 'Debloq Consigne'
   Rectangle "Rectangle_43" at 204,549 size 20x20
      Appearance <- "Var_Convoyeur_Carton_ConvoyeurC03_AcquitDefaut"
   TextField "Champ de texte_44" at 230,547 size 134x25; Text 'Acquit defaut'
   TextField "Champ de texte_45" at 230,461 size 158x25; Text 'Debloq fonction'
   IOField "Champ d'E/S_1" at 212,607 size 109x32; FormatPattern s99999
      ProcessValue <- "Var_Convoyeur_Carton_ConvoyeurC03_Consigne"
   TextField "Champ de texte_46" at 216,582 size 92x25; Text 'Consigne'
   Rectangle "Rectangle_11" at 590,217 size 20x20
      Appearance <- "Var_Convoyeur_Carton_ConvoyeurC03_EcartVitesse"
   TextField "Champ de texte_10" at 616,215 size 127x25; Text 'Ecart Vitesse'
   Rectangle "Rectangle_12" at 590,239 size 20x20
      Appearance <- "Var_Convoyeur_Carton_ConvoyeurC03_CommandeDemander"
   TextField "Champ de texte_11" at 616,237 size 212x25; Text 'Commande demandée'
   Rectangle "Rectangle_13" at 590,261 size 20x20
      Appearance <- "Var_Convoyeur_Carton_ConvoyeurC03_VitesseMaxAtteinte"
   TextField "Champ de texte_12" at 616,259 size 199x25; Text 'Vitesse max atteinte'
   Rectangle "Rectangle_14" at 590,283 size 20x20
      Appearance <- "Var_Convoyeur_Carton_ConvoyeurC03_Limite"
   TextField "Champ de texte_13" at 616,281 size 182x25; Text 'Limites de courant'
   Rectangle "Rectangle_15" at 590,305 size 20x20
      Appearance <- "Var_Convoyeur_Carton_ConvoyeurC03_FreinMoteur"
   TextField "Champ de texte_14" at 616,303 size 126x25; Text 'Frein Moteur'
   Rectangle "Rectangle_16" at 590,327 size 20x20
      Appearance <- "Var_Convoyeur_Carton_ConvoyeurC03_AlarmeSurchauffe"
   TextField "Champ de texte_15" at 616,325 size 181x25; Text 'Alarme Surchauffe'
   Rectangle "Rectangle_17" at 590,349 size 20x20
      Appearance <- "Var_Convoyeur_Carton_ConvoyeurC03_MoteurSensAvant"
   TextField "Champ de texte_16" at 616,347 size 180x25; Text 'Moteur sens avant'
   Rectangle "Rectangle_18" at 590,371 size 20x20
      Appearance <- "Var_Convoyeur_Carton_ConvoyeurC03_SurchargeMoteur"
   TextField "Champ de texte_17" at 616,369 size 174x25; Text 'Surcharge Moteur'
   TextField "Champ de texte_18" at 571,146 size 347x25; Text 'SORTIES'
   TextField "Champ de texte_19" at 590,192 size 85x25; Text '%ID264'
   Rectangle "Rectangle_20" at 590,394 size 20x20
      Appearance <- "Var_Convoyeur_Carton_ConvoyeurC03_PretEnclenchement"
   TextField "Champ de texte_20" at 616,392 size 193x25; Text 'Pret enclenchement'
   Rectangle "Rectangle_21" at 590,416 size 20x20
      Appearance <- "Var_Convoyeur_Carton_ConvoyeurC03_PretFonctionnement"
   TextField "Champ de texte_21" at 616,414 size 210x25; Text 'Pret Fonctionnement'
   Rectangle "Rectangle_22" at 590,438 size 20x20
      Appearance <- "Var_Convoyeur_Carton_ConvoyeurC03_Fonctionnement_Debloq"
   TextField "Champ de texte_22" at 616,436 size 236x25; Text 'Fonctionnement debloq.'
   Rectangle "Rectangle_23" at 590,460 size 20x20
      Appearance <- "Var_Convoyeur_Carton_ConvoyeurC03_DefautActif"
   Rectangle "Rectangle_24" at 590,482 size 20x20
      Appearance <- "Var_Convoyeur_Carton_ConvoyeurC03_Arret2Etat"
   TextField "Champ de texte_23" at 616,480 size 138x25; Text 'Arret 2 inactif'
   Rectangle "Rectangle_25" at 590,504 size 20x20
      Appearance <- "Var_Convoyeur_Carton_ConvoyeurC03_Arret3Etat"
   TextField "Champ de texte_24" at 616,502 size 138x25; Text 'Arret 3 inactif'
   Rectangle "Rectangle_26" at 590,526 size 20x20
      Appearance <- "Var_Convoyeur_Carton_ConvoyeurC03_BlocageActif"
   TextField "Champ de texte_25" at 616,524 size 135x25; Text 'Blocage actif'
   Rectangle "Rectangle_27" at 590,548 size 20x20
      Appearance <- "Var_Convoyeur_Carton_ConvoyeurC03_AlarmeActive"
   TextField "Champ de texte_26" at 616,546 size 134x25; Text 'Alarme active'
   TextField "Champ de texte_27" at 616,460 size 118x25; Text 'Défaut actif'
   IOField "Champ d'E/S_2" at 598,606 size 96x32; FormatPattern s99999
      ProcessValue <- "Var_Convoyeur_Carton_ConvoyeurC03_Vitesse"
   TextField "Champ de texte_28" at 602,581 size 73x25; Text 'Vitesse'
   Button "Bouton_1" at 8,8 size 96x32; TextOff 'Text'
   Button "Bouton_2" at 26,386 size 140x53; TextOff 'Convoyeur 01'
      on Release: ActivateScreen("Visu_ES_Variateur_C1", 0)
   Button "Bouton_3" at 25,450 size 140x53; TextOff 'Convoyeur 02'
      on Release: ActivateScreen("Visu_ES_Variateur_C2", 0)
   Button "Bouton_4" at 25,514 size 140x53; TextOff 'Convoyeur 03'
      on Release: ActivateScreen("Visu_ES_Variateur_C3", 0)

screen "TP_Robots" 1280x800, template "Modèle_1"
   Button "Bouton_1" at 37,399 size 159x95; TextOff 'Depart Cycle TP'
      on Release: ResetBit("Bits_B_Dcy")
      on Press: SetBit("Bits_B_Dcy")
      Appearance <- "B_VOY_DCY"
   Button "Bouton_2" at 37,496 size 158x86; TextOff 'Arret Cycle TP'
      on Release: ResetBit("Bits_B_Acy")
      on Press: SetBit("Bits_B_Acy")
      Appearance <- "B_VOY_ACY"
   GraphicView "Vue de graphique_3" at 230,144 size 1023x553; Picture "Capture d’écran 2023-07-10 135110"
   TextField "Champ de texte_1" at 31,140 size 158x25; Text 'CDT DE MARCHE'
   Rectangle "Rectangle_8" at 29,183 size 24x24
      Appearance <- "I_En_Arret_Urgence"
   TextField "Champ de texte_2" at 55,184 size 143x25; Text 'Arret Urgence'
   Rectangle "Rectangle_9" at 29,211 size 24x24
      Appearance <- "I_En_Automatique"
   TextField "Champ de texte_3" at 55,212 size 113x25; Text 'Mode Auto'
   Rectangle "Rectangle_10" at 29,239 size 24x24
      Appearance <- "I_En_Service"
   TextField "Champ de texte_4" at 61,240 size 103x25; Text 'En Service'
   Button "Bouton_3" at 1177,723 size 96x70; TextOff 'IN / OUT'
      on Release: ActivateScreen("Visu_ES-Cpu", 0)
   Button "Bouton_4" at 95,721 size 96x70; TextOff 'Alarmes'
      on Release: ActivateScreen("Alarmes", 0)
      Appearance <- "Bits_B_defaut_en_cours"
   GraphicView "Vue de graphique_5" at 19,728 size 60x60; Picture "Graphique_1"
      Visibility <- "Bits_B_defaut_en_cours"
   Button "Bouton_5" at 1070,723 size 96x70; TextOff 'PARAM'
      on Release: ActivateScreen("Parametrage", 0)
   Button "Bouton_7" at 856,723 size 96x70; TextOff 'TP Robots'
      Appearance <- "B_Pret_TP_Robotique"
      on Release: InvertBit("Bits_B_TP_Robot"); ResetBit("Bits_B_Demo_Hyppo")
   Button "Bouton_8" at 749,723 size 96x70; TextOff 'INIT.'
      on Release: ResetBit("Touche_Tch_Init")
      on Press: SetBit("Touche_Tch_Init")
   Button "Bouton_9" at 642,723 size 96x70; TextOff 'DEMO. HIPPO'
      on Release: InvertBit("Bits_B_Demo_Hyppo"); ResetBit("Bits_B_TP_Robot"); ActivateScreen("Principale", 0)
      Appearance <- "Bits_Pret_Demo_Hippo"
   Button "Bouton_10" at 535,723 size 96x70; TextOff 'Text'
   Button "Bouton_11" at 428,723 size 96x70; TextOff 'Text'
   Button "Bouton_12" at 321,723 size 96x70; TextOff 'HOME'
      on Click: ActivateScreen("Principale", 0)
   Button "Bouton_13" at 214,723 size 96x70; TextOff 'Acquit Defaut'
      on Release: ResetBit("Touche_Tch_Acquit")
      on Press: SetBit("Touche_Tch_Acquit")
   Circle "Cercle_1" at 473,447 size 28x28
      Visibility <- "Défauts_Defauts{0}"
      Appearance <- "Défauts_Defauts{0}"
   Circle "Cercle_2" at 358,447 size 28x28
      Visibility <- "Défauts_Defauts{1}"
      Appearance <- "Défauts_Defauts{1}"
   Circle "Cercle_3" at 266,512 size 28x28
      Visibility <- "Défauts_Defauts{2}"
      Appearance <- "Défauts_Defauts{2}"
   Circle "Cercle_4" at 412,565 size 28x28
      Visibility <- "Défauts_Defauts{12}"
      Appearance <- "Défauts_Defauts{12}"
   Circle "Cercle_5" at 629,564 size 28x28
      Visibility <- "Défauts_Defauts{13}"
      Appearance <- "Défauts_Defauts{13}"
   Circle "Cercle_6" at 760,504 size 28x28
      Visibility <- "Défauts_Defauts{14}"
      Appearance <- "Défauts_Defauts{14}"
   Circle "Cercle_7" at 615,447 size 28x28
      Visibility <- "Défauts_Defauts{15}"
      Appearance <- "Défauts_Defauts{15}"
   Circle "Cercle_8" at 775,565 size 28x28
      Visibility <- "Défauts_Defauts{3}"
      Appearance <- "Défauts_Defauts{3}"
   Circle "Cercle_9" at 760,437 size 28x28
      Visibility <- "Défauts_Defauts{4}"
      Appearance <- "Défauts_Defauts{4}"
   Circle "Cercle_10" at 262,447 size 28x28
      Visibility <- "Défauts_Defauts{5}"
      Appearance <- "Défauts_Defauts{5}"
   Circle "Cercle_11" at 262,571 size 28x28
      Visibility <- "Défauts_Defauts{6}"
      Appearance <- "Défauts_Defauts{6}"
   Circle "Cercle_12" at 963,392 size 28x28
      Visibility <- "Défauts_Defauts{7}"
      Appearance <- "Défauts_Defauts{7}"
   Circle "Cercle_13" at 1096,276 size 28x28
      Visibility <- "Défauts_Defauts{16}"
      Appearance <- "Défauts_Defauts{16}"
   Circle "Cercle_14" at 904,284 size 28x28
      Visibility <- "Défauts_Defauts{17}"
      Appearance <- "Défauts_Defauts{17}"
   Circle "Cercle_15" at 862,447 size 28x28
      Visibility <- "Défauts_Defauts{8}"
      Appearance <- "Défauts_Defauts{8}"
   Circle "Cercle_16" at 861,416 size 28x28
      Visibility <- "Défauts_Defauts{9}"
      Appearance <- "Défauts_Defauts{9}"
   Circle "Cercle_17" at 931,447 size 28x28
      Visibility <- "Défauts_Defauts{11}"
      Appearance <- "Défauts_Defauts{11}"
   Circle "Cercle_18" at 931,416 size 28x28
      Visibility <- "Défauts_Defauts{10}"
      Appearance <- "Défauts_Defauts{10}"
   Circle "Cercle_19" at 683,495 size 28x28
      Visibility <- "Défauts_Defauts{20}"
      Appearance <- "Défauts_Defauts{20}"
   Circle "Cercle_20" at 989,534 size 28x28
      Visibility <- "Défauts_Defauts{21}"
      Appearance <- "Défauts_Defauts{21}"
   Circle "Cercle_21" at 1050,284 size 28x28
      Visibility <- "Défauts_Defauts{22}"
      Appearance <- "Défauts_Defauts{22}"
   Circle "Cercle_22" at 1059,160 size 28x28
      Visibility <- "Défauts_Defauts{23}"
      Appearance <- "Défauts_Defauts{23}"
   Circle "Cercle_23" at 721,379 size 28x28
      Visibility <- "Défauts_Defauts{24}"
      Appearance <- "Défauts_Defauts{24}"
   Circle "Cercle_24" at 262,513 size 28x28
      Visibility <- "Défauts_Defauts{25}"
      Appearance <- "Défauts_Defauts{25}"
   Rectangle "Rectangle_1" at 825,454 size 20x20
      Appearance <- "I_det_Phot_01"
   Rectangle "Rectangle_2" at 975,454 size 20x20
      Appearance <- "I_det_Phot_02"
   Rectangle "Rectangle_3" at 1124,454 size 20x20
      Appearance <- "I_det_Phot_03"
   Rectangle "Rectangle_4" at 957,344 size 20x20
      Appearance <- "I_Det_Photo_7"
   Rectangle "Rectangle_12" at 862,344 size 20x20
      Appearance <- "I_Det_Photo_8"
   Rectangle "Rectangle_13" at 779,344 size 20x20
      Appearance <- "I_Det_Photo_9"
   Rectangle "Rectangle_14" at 1169,168 size 20x20
      Appearance <- "I_det_photo_03"
   Rectangle "Rectangle_15" at 1260,0 size 20x20
      Appearance <- "I_Det_Photo_9"
   Rectangle "Rectangle_16" at 1169,270 size 20x20
      Appearance <- "I_det_photo_02"
   Rectangle "Rectangle_17" at 1169,372 size 20x20
      Appearance <- "I_det_photo_01"
   Circle "Cercle_25" at 348,499 size 28x28
      Visibility <- "Défauts_Defauts{26}"
      Appearance <- "Défauts_Defauts{26}"
   Rectangle "Rectangle_18" at 29,267 size 24x24
      Appearance <- "I_Wieland_Au_porte01"
   TextField "Champ de texte_5" at 61,267 size 155x25; Text 'Porte Ouverte 1'
   Rectangle "Rectangle_19" at 29,295 size 24x24
      Appearance <- "I_Wieland_Au_Porte02"
   TextField "Champ de texte_6" at 61,295 size 155x25; Text 'Porte Ouverte 2'
   Rectangle "Rectangle_20" at 29,323 size 24x24
      Appearance <- "I_Wieland_Porte_non_Réarmée"
   TextField "Champ de texte_7" at 61,323 size 144x25; Text 'Porte Réarmée'
   TextField "Champ de texte_8" at 616,424 size 29x25; Text '01'
   TextField "Champ de texte_9" at 474,424 size 29x25; Text '02'
   TextField "Champ de texte_10" at 357,424 size 29x25; Text '03'
   TextField "Champ de texte_11" at 219,514 size 29x25; Text '04'
   TextField "Champ de texte_12" at 411,594 size 29x25; Text '05'
   TextField "Champ de texte_13" at 628,592 size 29x25; Text '06'
   TextField "Champ de texte_14" at 789,505 size 29x25; Text '07'
   Button "Bouton_14" at 4,5 size 124x122; TextOff 'Text'
      on Click: ActivateScreen("Page_demarrage", 0)
   TextField "Champ de texte_15" at 31,630 size 170x46; Text 'INITIALISATION EN COURS'
      Visibility <- "Bits_B_dmd_Init_robot"
      Appearance <- "Bits_B_dmd_Init_robot"
   TextField "Text field_1" at 331,163 size 404x81; Text 'TP_ROBOTS'
   Button "Bouton_15" at 963,723 size 96x70; TextOff 'MODE MANUEL'
      on Release: ActivateScreen("Mode_Manuel_B01_std_1", 0)
      Appearance <- "Bits_Globaux_x_En_manu"
      ObjectEnable <- "Bits_Globaux_x_En_manu"

screen "Visu_ES-Fanuc" 1280x800, template "Modèle_ES"
   GraphicView "Vue de graphique_1" at 24,140 size 272x158; Picture "Graphique_3"
   Rectangle "Rectangle_1" at 338,213 size 20x20
      Appearance <- "Fanuc1_Auto"
   TextField "Champ de texte_1" at 364,211 size 105x25; Text 'Mode auto'
   Rectangle "Rectangle_9" at 548,213 size 20x20
      Appearance <- "Fanuc2_Auto"
   TextField "Champ de texte_9" at 574,211 size 107x25; Text 'Mode Auto'
   TextField "Champ de texte_33" at 319,142 size 459x25; Text 'ENTREES'
   TextField "Champ de texte_34" at 338,188 size 91x25; Text 'Fanuc 01'
   TextField "Champ de texte_36" at 548,188 size 91x25; Text 'Fanuc 02'
   Rectangle "Rectangle_36" at 813,213 size 20x20
      Appearance <- "Fanuc1_Autor_Prise"
   TextField "Champ de texte_38" at 839,211 size 117x25; Text 'Autor_Prise'
   Rectangle "Rectangle_37" at 813,235 size 20x20
      Appearance <- "Fanuc1_Autor_vers_Fanuc02"
   TextField "Champ de texte_39" at 839,233 size 202x25; Text 'Autor_vers_Fanuc02'
   Rectangle "Rectangle_44" at 1023,213 size 20x20
      Appearance <- "Fanuc2_Autor_Prise"
   TextField "Champ de texte_46" at 1049,211 size 117x25; Text 'Autor_Prise'
   Rectangle "Rectangle_45" at 1023,235 size 20x20
      Appearance <- "Fanuc2_Autor_Depose"
   TextField "Champ de texte_47" at 1049,233 size 140x25; Text 'Autor_Depose'
   TextField "Champ de texte_70" at 794,142 size 459x25; Text 'SORTIES'
   TextField "Champ de texte_71" at 813,188 size 91x25; Text 'Fanuc 01'
   TextField "Champ de texte_73" at 1023,188 size 91x25; Text 'Fanuc 02'

screen "Mode_Manuel_Vision" 1280x800, template "Modèle_Manu"
   TextField "Champ de texte_34" at 35,138 size 584x25; Text 'Vision'
   Button "Bouton_1" at 39,179 size 169x68; TextOff 'Envoi trigger'
      on Release: ResetBit("Touche_Tch_Manu{92}")
      on Press: SetBit("Touche_Tch_Manu{92}")
      Appearance <- "O_Rentrer_Butée_01"
   Button "Bouton_2" at 226,179 size 245x71; TextOff 'x_Prise_disponible_UR'
      on Press: function_b14e0dd5("Touche_Tch_Manu{93}", 0)
      Appearance <- "O_Rentrer_Butée_01"
   TextField "Champ de texte_15" at 639,140 size 584x25; Text 'Porte Poste Vision'
   Button "Bouton_19" at 643,181 size 169x68; TextOff 'OUVRIR PORTE'
      on Press: function_b14e0dd5("32_Cmd_porte_vision_DB_x_Ouverture_porte_manu", 0)
   Button "Bouton_21" at 824,181 size 169x68; TextOff 'FERMER PORTE'
      on Press: function_b14e0dd5("32_Cmd_porte_vision_DB_x_Fermeture_porte_manu", 0)
   Rectangle "Rectangle_19" at 1008,183 size 20x20
      Appearance <- "I_porte_vision_op"
   TextField "Champ de texte_16" at 1034,181 size 137x25; Text 'Porte Ouverte'
   Rectangle "Rectangle_20" at 1008,205 size 20x20
      Appearance <- "I_porte_vision_cl"
   TextField "Champ de texte_17" at 1034,203 size 131x25; Text 'Porte Fermée'
   Rectangle "Rectangle_37" at 1008,235 size 20x20
      Appearance <- "O_Op_Porte_Vision"
   TextField "Champ de texte_32" at 1034,233 size 121x25; Text 'Ouvrir Porte'
   Rectangle "Rectangle_38" at 1008,257 size 20x20
      Appearance <- "O_Cl_porte_Vision"
   TextField "Champ de texte_33" at 1034,255 size 128x25; Text 'Fermer Porte'

screen "Mode_Manuel_B01_std_2" 1280x800, template "Modèle_Manu"
   ScreenModuleView "Poste Hippodrome_1" at 66,131 size 518x287; ScreenModuleType ""
      Guid_{11997190-69173} <- "DB_Stations_Station{5}"
   ScreenModuleView "Poste Hippodrome_2" at 623,133 size 518x287; ScreenModuleType ""
      Guid_{11997190-69173} <- "DB_Stations_Station{6}"
   ScreenModuleView "Poste Hippodrome_3" at 67,425 size 518x287; ScreenModuleType ""
      Guid_{11997190-69173} <- "DB_Stations_Station{7}"

screen "Mode_Manuel_B01_std_1" 1280x800, template "Modèle_Manu"
   ScreenModuleView "Poste Hippodrome_1" at 66,131 size 518x287; ScreenModuleType ""
      Guid_{11997190-69173} <- "DB_Stations_Station{1}"
   ScreenModuleView "Poste Hippodrome_2" at 623,133 size 518x287; ScreenModuleType ""
      Guid_{11997190-69173} <- "DB_Stations_Station{2}"
   ScreenModuleView "Poste Hippodrome_3" at 67,425 size 518x287; ScreenModuleType ""
      Guid_{11997190-69173} <- "DB_Stations_Station{3}"
   ScreenModuleView "Poste Hippodrome_4" at 624,427 size 518x287; ScreenModuleType ""
      Guid_{11997190-69173} <- "DB_Stations_Station{4}"

screen "Mode_Manuel_Imprimantes" 1280x800, template "Modèle_Manu"
   ScreenModuleView "Etat_imprimante_3D_1" at 31,135 size 397x275; ScreenModuleType ""
      Guid_{11997190-72965} <- "DB_Imprimantes_Imprimante{1}"
   ScreenModuleView "Etat_imprimante_3D_2" at 437,135 size 397x275; ScreenModuleType ""
      Guid_{11997190-72965} <- "DB_Imprimantes_Imprimante{2}"
   ScreenModuleView "Etat_imprimante_3D_3" at 843,135 size 397x275; ScreenModuleType ""
      Guid_{11997190-72965} <- "DB_Imprimantes_Imprimante{3}"
   ScreenModuleView "Etat_imprimante_3D_4" at 31,427 size 397x275; ScreenModuleType ""
      Guid_{11997190-72965} <- "DB_Imprimantes_Imprimante{4}"

PopupScreen "PopUp_Imp3d_1" 410x290
   ScreenModuleView "Etat_imprimante_3D_1" at 8,7 size 397x275; ScreenModuleType ""
      Guid_{11997190-72965} <- "DB_Imprimantes_Imprimante{1}"

PopupScreen "PopUp_Imp3d_2" 410x290
   ScreenModuleView "Etat_imprimante_3D_1" at 8,7 size 397x275; ScreenModuleType ""
      Guid_{11997190-72965} <- "DB_Imprimantes_Imprimante{2}"

PopupScreen "PopUp_Imp3d_3" 410x290
   ScreenModuleView "Etat_imprimante_3D_1" at 8,7 size 397x275; ScreenModuleType ""
      Guid_{11997190-72965} <- "DB_Imprimantes_Imprimante{3}"

PopupScreen "PopUp_Imp3d_4" 410x290
   ScreenModuleView "Etat_imprimante_3D_1" at 8,7 size 397x275; ScreenModuleType ""
      Guid_{11997190-72965} <- "DB_Imprimantes_Imprimante{4}"

